(* Logix 5000 project; controller TFF vendor 1 type 14 code 107 rev 33.11; software revision 33.04; part 14 of 38 *)
(* tags used below, declared in another part *)
   ActionCode : DINT;   // Action Code
   ActionProperty : DINT;   // Action Property
   ActionStructure : DINT;   // Action Data Structure
   ActionTag : DINT;   // Action Tag
   ActionValue : REAL;   // Action Value
   Boolean : DINT;   // Boolean Operator
   Branch : BOOL;   // Conditional Branch Flag
   BranchStep : DINT;   // Branch Step Number
   BufferStep : DINT;   // Buffer Step
   Clear : BOOL;   // Clear Operation Table Flag
   Code : DINT;   // Global Code
   Criteria1BoolValue : BOOL;   // Criteria 1 Discrete Value
   Criteria1Code : DINT;   // Criteria 1 Code
   Criteria1Met : BOOL;   // Criteria 1 Met
   Criteria1Operator : DINT;   // Criteria 1 Operator
   Criteria1Property : DINT;   // Criteria 1 Property
   Criteria1RealValue : REAL;   // Criteria 1 Real Value
   Criteria1Structure : DINT;   // Criteria 1 Data Structure
   Criteria1Tag : DINT;   // Criteria 1 Tag
   Criteria1Type : BOOL;   // Criteria 1 Type 0=Real, 1=Boolean
   Criteria1Value : REAL;   // Criteria 1 Value
   Criteria2BoolValue : BOOL;   // Criteria 2 Discrete Value
   Criteria2Code : DINT;   // Criteria 2 Code
   Criteria2Met : BOOL;   // Criteria 2 Met
   Criteria2Operator : DINT;   // Criteria 2 Operator
   Criteria2Property : DINT;   // Criteria 2 Property
   Criteria2RealValue : REAL;   // Criteria 2 Real Value
   Criteria2Structure : DINT;   // Criteria 2 Data Structure
   Criteria2Tag : DINT;   // Criteria 2 Tag
   Criteria2Type : BOOL;   // Criteria 2 Type 0=Real, 1=Boolean
   Criteria2Value : REAL;   // Criteria 2 Value
   CriteriaMet : BOOL;   // Criteria Met
   DateTime : DINT[7];   // Date and Time
   ErrorCheck : BOOL;   // Error Check Flag
   Index : DINT;   // Index
   LastStep : DINT;   // Last Step
   NextStep : DINT;   // Next Step
   PendingStep : DINT;   // Current Step
   PhaseClear : BOOL;   // Phase Clear
   PhaseClearNumber : DINT;   // Phase Clear Number
   PhaseNumber : DINT;   // Phase FOR NEXT Index
   Pointer : DINT;   // Pointer
   PreRunLog : BOOL;   // Log Pre Run Set Points
   Property : DINT;   // Case Property
   Run : BOOL;   // Operation Run Status
   sAction : STRING10;   // Action Code String
   sActionProperty : STRING4;   // Action Property String
   sActionStructure : STRING4;   // Action Data Structure String
   sActionTag : STRING4;   // Action Tag String
   sBufferEvents : STRING50;   // Buffer Events String
   sCode : STRING10;   // Global code String
   sColon : STRING4;   // Colon separator String
   sComma : STRING4;   // Comma String
   sCriteria1 : STRING10;   // Criteria 1 Code String
   sCriteria1Property : STRING4;   // Criteria 1 Property String
   sCriteria1Structure : STRING4;   // Criteria 1 Data Structure String
   sCriteria1Tag : STRING4;   // Criteria 1 Tag String
   sCriteria2 : STRING10;   // Criteria 2 Code String
   sCriteria2Property : STRING4;   // Criteria 2 Property String
   sCriteria2Structure : STRING4;   // Criteria 2 Data Structure String
   sCriteria2Tag : STRING4;   // Criteria 2 Tag String
   sDateTime : STRING25;   // Date and Time String
   sPeriod : STRING4;   // Timer separator String
   sProperty : STRING4;   // Property String
   sStructure : STRING4;   // Structure String
   sTag : STRING4;   // Tag String
   sTemp : STRING50;   // Temp String
   Structure : DINT;   // Structure code
   sZero : STRING4;   // Zero String
   Tag : DINT;   // Tag value
   TempEvents : DINT;   // Temp Register
   TempSteps : DINT;
   Tenths : DINT;   // Thents (Date and Time management)
   ThisStep : DINT;   // This Step (Error management)
   Value : REAL;   // Temp Value
   AlarmAnalog : AlarmAnalog[50];   // Analog Alarm Array
   AlarmControl : AlarmControl;   // Alarm Control
   AlarmDeviation : AlarmDeviation[20];   // Control Loop Deviation Alarm Array
   AnalogPoint : AnalogInput[50];   // Analog Input Array
   BagInflate : BagInflate;
   CCPSystem : CCPSystem;   // CCP System Data
   ChartMark : ChartMark;   // Chart Mark
   Concentration : Concentration;
   ControlLoop : ControlLoop[20];   // Control Loop Array
   CPU_Scanning : BOOL;   // System Scanning Flag
   CriteriaFlag : CriteriaFlag;   // Criteria Flag used in CCP Recipe
   DerivedData : DerivedData;   // Derived data (user input and calculated values)
   Diafiltration : Diafiltration;
   DigitalPoint : DigitalPoint[150];   // Digital Point Array
   Drive : Drive[11];   // Drives Array
   Exchange_OUT : Exchange_OUT;   // Exchange Outputs
   ExternalTCU : BOOL;   // Use of External TCU
   ExternalWeight : BOOL;   // Use of External Weight
   FirstScanComplete : BOOL;   // First Scan Complete Flag
   FlowPath : FlowPath[64];   // Flow Path Array
   FQ_Conc : ALIAS FOR Totalizer[0];   // Concentration Totalizer
   FQ_Diaf : ALIAS FOR Totalizer[1];   // DiafiltrationTotalizer
   Gateway : Gateway;   // Gateway Control
   HoldTime : ALIAS FOR Timers[20];   // Hold Time
   LogVal : LoggedValue;   // Setpoints to be logged
   Membrane_Data : Membrane_Data;   // Membrane Data
   MiscBOOL : BOOL[64];   // Misc BOOL Values
   MiscDINT : DINT[32];   // Misc DINT Values
   MiscREAL : REAL[50];   // Misc Real Values
   Mixer : Mixer;   // Mixer config. structure
   Operation : Operation[6,251];   // Operation Table
   PCV101_Control : PCV_Control;   // PCV101 Control UDT
   PCV201_Control : PCV_Control;   // PCV201 Control UDT
   Phase : Phases[6];   // Phase Control Array
   Phase0 : ALIAS FOR Phase[0];   // Phase 0
   Phase0_Totalizer_Feed : ALIAS FOR PhaseTotalizer[0];   // Phase 0 Total Feed
   Phase0_Totalizer_Filtrate : ALIAS FOR PhaseTotalizer[6];   // Phase 0 Total Filtrate
   Phase0_Totalizer_Transfer : ALIAS FOR PhaseTotalizer[12];   // Phase 0 Total Transfer
   Phase1 : ALIAS FOR Phase[1];   // Phase 1
   Phase2 : ALIAS FOR Phase[2];   // Phase 2
   Phase3 : ALIAS FOR Phase[3];   // Phase 3
   Phase4 : ALIAS FOR Phase[4];   // Phase 4
   Phase5 : ALIAS FOR Phase[5];   // Phase 5
   PhaseTotalizer : PhaseTotalizer[18];   // Phase Totalizers Array
   PLCFault : FaultRecordType;   // PLC Major Fault Record
   ProcedureTime : ALIAS FOR Timers[19];   // Procedure Time
   Prompt : Prompt[7];   // Prompt Array
   Prompt0 : ALIAS FOR Prompt[0];   // Phase 0 Prompt
   Prompt1 : ALIAS FOR Prompt[1];   // Phase 1 Prompt
   Prompt2 : ALIAS FOR Prompt[2];   // Phase 2 Prompt
   Prompt3 : ALIAS FOR Prompt[3];   // Phase 3 Prompt
   Prompt4 : ALIAS FOR Prompt[4];   // Phase 4 Prompt
   Prompt5 : ALIAS FOR Prompt[5];   // Phase 5 Prompt
   SysControl : SysControl;   // General system status and command
   ThisSystem : SystemType;
   TIC101Control : TCUControl;
   TimerControl : TimerControl;   // Timer Control
   Timers : Timers[22];   // Timer Array
   Totalizer : Totalizers[20];   // Totalizers Array
   UserAlarm : UserAlarm;   // User Alarm (used in CCP Recipe)
   UserTotalizerManagement : UserTotalizerManagement;   // User Totalizer management
   Valve : Valve[100];   // Valve Array
   Y500A : ALIAS FOR DigitalOutput[10];
   Y500B : ALIAS FOR DigitalOutput[11];
   Y501A : ALIAS FOR DigitalOutput[12];
   Y501B : ALIAS FOR DigitalOutput[13];
   YA10 : ALIAS FOR DigitalPoint[59];
(* CCPSystem, continued *)

ROUTINE Branch   (* structured text *)
// Branch to Label Routine
   (* =======================================================================
   	Branch : Conditionnal branch management
   
   	List of treatments
   		- Get current action code
   		- Extract informations based on action code
   		- Jump to label and Jump Step processing
   
   -----------------------------------------------------------------------------------------------------------------------------------------------------
   	History
   		2019-DEC-24 - Merck - Q. Spindler - Initial version for Candidate Release 1.00.00.00.a
   =========================================================================*)
   
   
   (* Get current action code
   =========================================================================*)
   (*Get the pending step Action Code and Action Value from the operation array*)
   ActionCode := Operation[PhaseNumber,PendingStep].Action;
   ActionValue := Operation[PhaseNumber,PendingStep].ActionValue;
   
   (* Extract informations based on action code
   =========================================================================*)
   (*Extract the Structure, Tag and Property values from the action code. The action code is
   in the format SSTTTPP*)
   IF ActionCode <> 0 THEN;
   	DTOS (ActionCode, sAction);
   	IF sAction.LEN = 7 THEN;
   		MID (sAction, 2, 1, sActionStructure);
   		MID (sAction, 3, 3, sActionTag);
   		MID (sAction, 2, 6, sActionProperty);
   	ELSIF sAction.LEN = 6 THEN;
   		MID (sAction, 1, 1, sActionStructure);
   		MID (sAction, 3, 2, sActionTag);
   		MID (sAction, 2, 5, sActionProperty);
   	END_IF;
   	STOD (sActionStructure, ActionStructure);
   	STOD (sActionTag, ActionTag);
   	STOD (sActionProperty, ActionProperty);
   ELSE;
   	ActionStructure := 0;
   	ActionProperty := 0;
   END_IF;
   
   (* Jump to label and Jump Step processing
   =========================================================================*)
   (*Check to determine if action is a conditional branch, Structure=7 and Property=5*)
   BranchStep := 0;
   Phase[PhaseNumber].Label := 0;
   IF ActionStructure = 7 AND ActionProperty = 5  AND NOT Prompt[PhaseNumber].Pending THEN;
   	IF CriteriaMet THEN;
   		FOR BranchStep := 1 TO 250 DO;
   		(*If Jump to label action exist copy the label value in corresponding Phase label*)
   			IF Operation[PhaseNumber, BranchStep].Label = ActionValue THEN;
   				Phase[PhaseNumber].Label := ActionValue;
   				EXIT;
   			END_IF;
   		END_FOR;
   	ELSE;
   		(*Jump to BufferSteps routine and update Actual step number*)
   		JSR (BufferSteps);
   		Phase[PhaseNumber].ActualStep := (PendingStep + 1);
   	END_IF;
   
   ELSIF Phase[PhaseNumber].JumpPLC THEN;
   	FOR BranchStep := 1 TO 250 DO;
   		IF Operation[PhaseNumber, BranchStep].Step = Phase[PhaseNumber].JumpStep THEN;
   			Phase[PhaseNumber].ActualStep := BranchStep;
   			EXIT;
   		END_IF;
   	END_FOR;
   END_IF;
   
END_ROUTINE

ROUTINE BufferEvents   (* structured text *)
// Event Log Buffer Routine
   (* =======================================================================
   	Buffer Events : This routine scans all event code values defined in the event array downloaded by CCP6
   					If the value of the tag referenced by the code has changed from the last scan,the time stamp,
   					action code and new/old values are written to the buffer.
   					The buffer pointer used by CCP6 is updated after scanning all tags
   
   	Warning :		This code should not be modified without a control of change impact on the Recipe download check procedure of CCPRuntime.exe
   
   	List of treatments
   		- Get current action code
   		- Extract informations based on event code
   		- Navigate through the event categories
   		- Log Pre-run values
   		- Build event contents
   		- Reset flag and pointer
   
   -----------------------------------------------------------------------------------------------------------------------------------------------------
   	History
   		2019-DEC-24 - Merck - Q. Spindler - Initial version for Candidate Release 1.00.00.00.a
   		2020-MAR-30 - Merck - Q. Spindler - Modifications for Candidate Release 1.00.00.00.b
   					- Replace ActionProperty by Property for TIC
   					- Add SysControl.Zero_WI101_Cmd
   					- Add Valve.ZSOverride for valves limit switch alarms
   					- Add Gateway events
   		2020-SEP-18 - Merck - Q. Spindler - Modifications for Candidate Release 1.00.00.00.d
   					- Add ExternalWeight and ExternalTCU events
   		2022-JAN-21 - Merck - Q. Spindler - Modifications for Candidate Release 1.01.00.00.a
   					- Change resetting of sStructure in case of wrong code length by DTOS function
   		2022-SEP-21 - Actemium - J. Jaekel - Modifications for Candidate Release 1.01.00.01.a
   					- Add K and Q factor events
   =========================================================================*)
   
   
   (* Get the current pointer value
   =========================================================================*)
   STOD (CCPSystem.BufferEvents[0], Pointer);
   
   (* Extract informations based on event code
   =========================================================================*)
   (*Index through the event listing and get current value for each code*)
   (*The first element in the array is the array length*)
   FOR Index := 1 TO CCPSystem.EventList.Event[0] DO;
   
   	(*Extract the Structure, Tag and Property values from the code.  The code is in the format SSTTTPP*)
   	Code := CCPSystem.EventList.Event[Index];
   	DTOS (Code, sCode);
   
   		IF sCode.LEN = 7 THEN;
   			MID (sCode, 2, 1, sStructure);
   			MID (sCode, 3, 3, sTag);
   			MID (sCode, 2, 6, sProperty);
   		ELSIF sCode.LEN = 6 THEN;
   			MID (sCode, 1, 1, sStructure);
   			MID (sCode, 3, 2, sTag);
   			MID (sCode, 2, 5, sProperty);
   		ELSE;
   			(*Ignore if code length is not 6 or 7*)
   			DTOS (0, sStructure);
   		END_IF;
   		STOD (sStructure, Structure);
   		STOD (sTag, Tag);
   		STOD (sProperty, Property);
   
   	(* Tag:= 0; (*put in to handel error in congig files*)
   
   	Value := 0;
   
   (* Navigate through the event categories
   =========================================================================*)
   	(*Get the value based on the structure, tag and property*)
   	CASE	Structure OF
   		1: 	CASE	Property OF (*Analog Alarms*)
   			1:	IF AlarmAnalog[Tag].Override THEN Value := 1; ELSE Value := 0; END_IF;
   			2:	Value := AlarmAnalog[Tag].LOLO;
   			3:	Value := AlarmAnalog[Tag].LO;
   			4:	Value := AlarmAnalog[Tag].HI;
   			5:	Value := AlarmAnalog[Tag].HIHI;
   			6:	IF AlarmAnalog[Tag].LOLOAlarm THEN Value := 1; ELSE Value := 0; END_IF;
   			7:	IF AlarmAnalog[Tag].LOAlarm THEN Value := 1; ELSE Value := 0; END_IF;
   			8:	IF AlarmAnalog[Tag].HIAlarm THEN Value := 1; ELSE Value := 0; END_IF;
   			9:	IF AlarmAnalog[Tag].HIHIAlarm THEN Value := 1; ELSE Value := 0; END_IF;
   			END_CASE;
   		2: 	CASE	Property OF (*Deviation Alarms*)
   			1:	IF AlarmDeviation[Tag].Override THEN Value := 1; ELSE Value := 0; END_IF;
   			4:	Value := AlarmDeviation[Tag].HI;
   			5:	Value := AlarmDeviation[Tag].HIHI;
   			8:	IF AlarmDeviation[Tag].HIAlarm THEN Value := 1; ELSE Value := 0; END_IF;
   			9:	IF AlarmDeviation[Tag].HIHIAlarm THEN Value := 1; ELSE Value := 0; END_IF;
   			END_CASE;
   		3: 	CASE	Property OF (*Digital Alarms*)
   			1:	IF DigitalPoint[Tag].Override THEN Value := 1; ELSE Value := 0; END_IF;
   			6:	IF DigitalPoint[Tag].Alarm THEN Value := 1; ELSE Value := 0; END_IF;
   			7:	IF DigitalPoint[Tag].CurrentValue THEN Value := 1; ELSE Value := 0; END_IF;
   			END_CASE;
   		4: 	CASE	Property OF (*Analog Inputs*)
   			1:	Value := AnalogPoint[Tag].CurrentValue;
   			2:	Value := AnalogPoint[Tag].ScaledMin;
   			3:	Value := AnalogPoint[Tag].ScaledMax;
   			END_CASE;
   		5:	CASE	Property OF (*Control Loops*)
   			1:	IF ControlLoop[Tag].Manual THEN Value := 1; ELSE Value := 0; END_IF;
   			2:	IF ControlLoop[Tag].Auto1 THEN Value := 1; ELSE Value := 0; END_IF;
   			3:	IF ControlLoop[Tag].Auto2 THEN Value := 1; ELSE Value := 0; END_IF;
   			4:	IF ControlLoop[Tag].Auto3 THEN Value := 1; ELSE Value := 0; END_IF;
   			5:	IF ControlLoop[Tag].Auto4 THEN Value := 1; ELSE Value := 0; END_IF;
   			6:	Value := ControlLoop[Tag].SPManual;
   			7:	Value := ControlLoop[Tag].SPAuto1;
   			8:	Value := ControlLoop[Tag].SPAuto2;
   			9:	Value := ControlLoop[Tag].SPAuto3;
   			10:	Value := ControlLoop[Tag].SPAuto4;
   			11:	Value := ControlLoop[Tag].RampRate;
   			12:	Value := ControlLoop[Tag].Deadband;
   			13:	Value := ControlLoop[Tag].StableTime;
   			14:	Value := ControlLoop[Tag].KP[0];
   			15:	Value := ControlLoop[Tag].KI[0];
   			16:	Value := ControlLoop[Tag].KD[0];
   			17:	Value := ControlLoop[Tag].DB[0];
   			18:	Value := ControlLoop[Tag].KP[1];
   			19:	Value := ControlLoop[Tag].KI[1];
   			20:	Value := ControlLoop[Tag].KD[1];
   			21:	Value := ControlLoop[Tag].DB[1];
   			22:	Value := ControlLoop[Tag].KP[2];
   			23:	Value := ControlLoop[Tag].KI[2];
   			24:	Value := ControlLoop[Tag].KD[2];
   			25:	Value := ControlLoop[Tag].DB[2];
   			26:	IF ControlLoop[Tag].Stable THEN Value := 1; ELSE Value := 0; END_IF;
   			27:	IF ControlLoop[Tag].DBOK THEN Value := 1; ELSE Value := 0; END_IF;
   			28:	IF ControlLoop[Tag].RampStatus THEN Value := 1; ELSE Value := 0; END_IF;
   			END_CASE;
   		7:	CASE	Property OF (*Phase Control*)
   			1:	IF Phase[Tag].Run THEN Value := 1; ELSE Value := 0; END_IF;
   			2:	IF Phase[Tag].Stop THEN Value := 1; ELSE Value := 0; END_IF;
   			3:	IF Phase[Tag].Hold THEN Value := 1; ELSE Value := 0; END_IF;
   			4:	IF Phase[Tag].Pause THEN Value := 1; ELSE Value := 0; END_IF;
   			5:	IF Phase[Tag].Label = 0 THEN CCPSystem.EventList.Value[Index] := 0; END_IF; (*Ignore change to 0*)
   				Value := Phase[Tag].Label;
   			6:	IF Phase[Tag].JumpPLC THEN Value := 1; ELSE Value := 0; END_IF;
   			END_CASE;
   		8: 	CASE	Property OF (*Prompts*)
   			1:	IF Prompt[Tag].PromptOK THEN Value := 1; ELSE Value := 0; END_IF;
   			2:	IF Prompt[Tag].PromptYesNO THEN Value := 1; ELSE Value := 0; END_IF;
   			3:	IF Prompt[Tag].ResponseOK THEN Value := 1; ELSE Value := 0; END_IF;
   			4:	IF Prompt[Tag].ResponseYes THEN Value := 1; ELSE Value := 0; END_IF;
   			5:	IF Prompt[Tag].ResponseNo THEN Value := 1; ELSE Value := 0; END_IF;
   			END_CASE;
   		9: 	CASE	Property OF (*Pumps*)
   			1:	IF Drive[Tag].RunStatus THEN Value := 1; ELSE Value := 0; END_IF;
   			2:	IF Drive[Tag].Direction THEN Value := 1;ELSE Value := 0; END_IF;
   			3:	IF Drive[Tag].Mode THEN Value := 1; ELSE Value := 0; END_IF;
   			END_CASE;
   		10:	CASE	Property OF (*Exchange Output*)
   			1:	Value := Exchange_OUT.AO01;
   			2:	Value := Exchange_OUT.AO02;
   			3:	Value := Exchange_OUT.AO03;
   			4:	Value := Exchange_OUT.AO04;
   			5:	IF Exchange_OUT.DO01 THEN Value := 1; ELSE Value := 0; END_IF;
   			6:	IF Exchange_OUT.DO02 THEN Value := 1; ELSE Value := 0; END_IF;
   			7:	IF Exchange_OUT.DO03 THEN Value := 1; ELSE Value := 0; END_IF;
   			8:	IF Exchange_OUT.DO04 THEN Value := 1; ELSE Value := 0; END_IF;
   			9:	IF Exchange_OUT.DO05 THEN Value := 1; ELSE Value := 0; END_IF;
   			10:	IF Exchange_OUT.DO06 THEN Value := 1; ELSE Value := 0; END_IF;
   			11:	IF Exchange_OUT.DO07 THEN Value := 1; ELSE Value := 0; END_IF;
   			12:	IF Exchange_OUT.DO08 THEN Value := 1; ELSE Value := 0; END_IF;
   			END_CASE;
   		11:	CASE	Property OF (*Timers*)
   			3:	IF Timers[Tag].Enable THEN Value := 1; ELSE Value := 0; END_IF;
   			4:	IF Timers[Tag].Reset THEN Value := 1; ELSE Value := 0; END_IF;
   			END_CASE;
   		13:	CASE	Property OF (*Valves*)
   			2:	Value := Valve[Tag].StatusWord;
   			3:	IF Valve[Tag].Mode THEN Value := 1; ELSE Value := 0; END_IF;
   			4:	IF Valve[Tag].Alarm THEN Value := 1; ELSE Value := 0; END_IF;
   			5:	Value := Valve[Tag].Status;
   			6:	IF Valve[Tag].ZSOverride THEN Value := 1; ELSE Value := 0; END_IF;
   			END_CASE;
   		14:	CASE	Property OF (*Agitator*)
   			1:	IF Mixer.Mode THEN Value := 1; ELSE Value := 0; END_IF;
   			2:	Value := Mixer.SPManual;
   			3:	Value := Mixer.SPAutoMin;
   			4:	Value := Mixer.SPAutoMax;
   			5:	Value := Mixer.LevelMin;
   			6:	Value := Mixer.LevelMax;
   			END_CASE;
   		15:	CASE	Property OF (*Misc.*)
   			1:	IF MiscBOOL[Tag] THEN Value := 1; ELSE Value := 0; END_IF;
   			2:	Value := MiscDINT[Tag];
   			3:	Value := MiscREAL[Tag];
   			END_CASE;
   		16:	CASE	Property OF (*Alarm Control*)
   			1:	IF AlarmControl.EnableAllOut THEN Value := 1; ELSE Value := 0; END_IF;
   			2:	IF AlarmControl.DisableAllOut THEN Value := 1; ELSE Value := 0; END_IF;
   			3:	IF AlarmControl.AckOutput THEN Value := 1; ELSE Value := 0; END_IF;
   			6:	IF AlarmControl.EnableAllAnaSigOut THEN Value := 1; ELSE Value := 0; END_IF;
   			7:	IF AlarmControl.DisableAllAnaSigOut THEN Value := 1; ELSE Value := 0; END_IF;
   			END_CASE;
   		17:	CASE	Property OF (*Miscellaneous*)
   			1:	IF SysControl.DefaultOut THEN Value := 1; ELSE Value := 0; END_IF;
   			2:	IF ChartMark.Out THEN Value := 1; ELSE Value := 0; END_IF;
   			3:	IF SysControl.AllAutoOut THEN Value := 1; ELSE Value := 0; END_IF;
   			4:	IF UserTotalizerManagement.LogUserOut THEN Value := 1; ELSE Value := 0; END_IF;
   			5:	IF UserTotalizerManagement.StartUser THEN Value := 1; ELSE Value := 0; END_IF;
   			6:	IF UserTotalizerManagement.ResetUserOut THEN Value := 1; ELSE Value := 0; END_IF;
   			7:	IF SysControl.Tare_WI101_Cmd THEN Value := 1; ELSE Value := 0; END_IF;
   			8:	IF SysControl.ClearTare_WI101_Cmd THEN Value := 1; ELSE Value := 0; END_IF;
   			9:	IF SysControl.UV_Auto_Zero_Cmd THEN Value := 1; ELSE Value := 0; END_IF;
   			10:	IF SysControl.Zero_WI101_Cmd THEN Value := 1; ELSE Value := 0; END_IF;
   			11:	IF CCPSystem.DefaultOnComplete THEN Value := 1; ELSE Value := 0; END_IF;
   			12:	IF UserAlarm.NonCritical1 THEN Value := 1; ELSE Value := 0; END_IF;
   			13:	IF UserAlarm.Critical1 THEN Value := 1; ELSE Value := 0; END_IF;
   			14:	IF UserAlarm.NonCritical2 THEN Value := 1; ELSE Value := 0; END_IF;
   			15:	IF UserAlarm.Critical2 THEN Value := 1; ELSE Value := 0; END_IF;
   			16:	IF SysControl.Tare_PI001_Cmd THEN Value := 1; ELSE Value := 0; END_IF;
   			17:	IF SysControl.Tare_PI101_Cmd THEN Value := 1; ELSE Value := 0; END_IF;
   			18:	IF SysControl.Tare_PI201_Cmd THEN Value := 1; ELSE Value := 0; END_IF;
   			19:	IF SysControl.Tare_PI401_Cmd THEN Value := 1; ELSE Value := 0; END_IF;
   			20:	IF SysControl.Tare_PI601_Cmd THEN Value := 1; ELSE Value := 0; END_IF;
   			21:	IF BagInflate.cmd THEN Value := 1; ELSE Value := 0; END_IF;
   			22:	IF ExternalTCU THEN Value := 1; ELSE Value := 0; END_IF;
   			23:	IF ExternalWeight THEN Value := 1; ELSE Value := 0; END_IF;
   			END_CASE;
   		18:	CASE	Property OF (*Criteria Flag*)
   			1:	IF CriteriaFlag.Flag1 THEN Value := 1; ELSE Value := 0; END_IF;
   			2:	IF CriteriaFlag.Flag2 THEN Value := 1; ELSE Value := 0; END_IF;
   			3:	IF CriteriaFlag.Flag3 THEN Value := 1; ELSE Value := 0; END_IF;
   			4:	IF CriteriaFlag.Flag4 THEN Value := 1; ELSE Value := 0; END_IF;
   			5:	IF CriteriaFlag.Flag5 THEN Value := 1; ELSE Value := 0; END_IF;
   			END_CASE;
   		19:	CASE	Property OF (*Concentration*)
   			1:	IF FQ_Conc.Enable THEN Value := 1; ELSE Value := 0; END_IF;
   			2:	IF FQ_Conc.Reset THEN Value := 1; ELSE Value := 0; END_IF;
   			3:	IF Concentration.LogConcOut THEN Value := 1; ELSE Value := 0; END_IF;
   			4:	Value := Concentration.Conc_Init ;
   			5:	Value := Concentration.Conc_Final ;
   			6:	Value := Concentration.Conc_Final_Volume ;
   			7:	Value := DerivedData.HOLDUP ;
   			10: IF Concentration.Final_Conc_Volume_Reached THEN Value := 1; ELSE Value := 0; END_IF;
   			11: IF Concentration.Final_Conc_Protein_Reached THEN Value := 1; ELSE Value := 0; END_IF;
   			END_CASE;
   		20:	CASE	Property OF (*Diafiltration*)
   			1:	IF FQ_Diaf.Enable THEN Value := 1; ELSE Value := 0; END_IF;
   			2:	IF FQ_Diaf.Reset THEN Value := 1; ELSE Value := 0; END_IF;
   			3:	IF Diafiltration.LogDiafOut THEN Value := 1; ELSE Value := 0; END_IF;
   			4:	IF Diafiltration.Snap THEN Value := 1; ELSE Value := 0; END_IF;
   			5:	Value := Diafiltration.Diaf_Init ;
   			6:	Value := Diafiltration.Diaf_Final_Volume ;
   			10: IF Diafiltration.Final_Diaf_Volum_Reached THEN Value := 1; ELSE Value := 0; END_IF;
   			END_CASE;
   		21:	CASE	Property OF (*Membrane Data*)
   			1:	Value := Membrane_Data.Area ;
   			2:	Value := Membrane_Data.Density ;
   			3:	Value := DerivedData.FI101Q ;
   			4:	Value := DerivedData.FI201Q ;
   			5:	Value := DerivedData.FI401Q ;
   			6:	Value := DerivedData.FI101K ;
   			7:	Value := DerivedData.FI201K ;
   			8:	Value := DerivedData.FI401K ;
   			END_CASE;
   		22:	CASE	Property OF (*Gateway*)
   			1:	IF Tag <=31 THEN; (*Digital Actions*)
   					IF Gateway.RecipeAction_Digital[0].[Tag] THEN	Value := 1; ELSE Value := 0; END_IF;
   				ELSIF Tag <=63 THEN;
   					IF Gateway.RecipeAction_Digital[1].[Tag-32] THEN	Value := 1; ELSE Value := 0; END_IF;
   				END_IF;
   			2:	IF Tag <=19 THEN; (*Analog Actions*)
   				Value := Gateway.RecipeAction_Analog[Tag];
   				END_IF;
   			END_CASE;
   		23:	CASE	Property OF (*PCV Control*)
   			1:	IF PCV101_Control.FullOpen THEN Value := 1; ELSE Value := 0; END_IF;
   			2:	IF PCV101_Control.FullClose THEN Value := 1; ELSE Value := 0; END_IF;
   			3:	IF PCV201_Control.FullOpen THEN Value := 1; ELSE Value := 0; END_IF;
   			4:	IF PCV201_Control.FullClose THEN Value := 1; ELSE Value := 0; END_IF;
   			END_CASE;
   		24:	CASE	Property OF (*Event value.*)
   			1:	Value := LogVal.Value[Tag];
   			END_CASE;
   		25: CASE	Property OF (*Flow Paths*)
   			1:	IF FlowPath[Tag].Status THEN Value := 1; ELSE Value := 0; END_IF;
   			END_CASE;
   		26: CASE	Property OF (*Clamshell*)
   			1:	IF Y500A THEN Value := 1; ELSE Value := 0; END_IF;
   			2:	IF Y500B THEN Value := 1; ELSE Value := 0; END_IF;
   			3:	IF Y501A THEN Value := 1; ELSE Value := 0; END_IF;
   			4:	IF Y501B THEN Value := 1; ELSE Value := 0; END_IF;
   			11:  IF ThisSystem.MoldType = 123 THEN Value := 1; ELSE Value := 0; END_IF;
   			12:  IF ThisSystem.MoldType = 124 THEN Value := 1; ELSE Value := 0; END_IF;
   			13:  IF ThisSystem.MoldType = 126 THEN Value := 1; ELSE Value := 0; END_IF;
   			21:  IF ThisSystem.PreviousValue = 123 THEN Value := 1; ELSE Value := 0; END_IF;
   			22:  IF ThisSystem.PreviousValue = 124 THEN Value := 1; ELSE Value := 0; END_IF;
   			23:  IF ThisSystem.PreviousValue = 126 THEN Value := 1; ELSE Value := 0; END_IF;
   			END_CASE;
   		27:	CASE	Property OF (*TIC*)
   				1:	IF TIC101Control.RunCommand THEN Value := 1; ELSE Value := 0; END_IF;
   				2:  IF TIC101Control.Mode THEN Value := 1; ELSE Value := 0; END_IF;
   				3:	Value := TIC101Control.Offset;
   				4:	Value := TIC101Control.OffsetTime;
   				5:	Value := TIC101Control.LevelMin;
   			END_CASE;
   	(*Missing else statement accepted for the purpose of proper integration with CCPRuntime.exe*)
   	END_CASE;
   
   (* Log Pre-run values
   =========================================================================*)
   	(*Record value for Pre-Run Log if flag is set*)
   	IF PreRunLog THEN;
   		CCPSystem.EventList.PreRunValue[Index] := Value;
   	END_IF;
   
   
   (* Build event contents
   =========================================================================*)
   	(*Check for change in value*)
   	IF CCPSystem.EventList.Value[Index] <> Value THEN;
   		(*Increment pointer*)
   		Pointer := Pointer + 1;
   		(*Roll over pointer if equal to max*)
   		IF Pointer = 251 THEN Pointer := 1; END_IF;
   
   		(*Concatenate the action code to the date/time and add comma*)
   		DTOS (Code, sTemp);
   		CONCAT(sDateTime, sTemp, sBufferEvents);
   		CONCAT(sBufferEvents, sComma, sBufferEvents);
   
   		(*Concatenate the new value and add comma*)
   		RTOS (Value, sTemp);
   		CONCAT (sBufferEvents, sTemp, sBufferEvents);
   		CONCAT (sBufferEvents, sComma, sBufferEvents);
   
   		(*Concatenate the old value and store in the buffer*)
   		RTOS(CCPSystem.EventList.Value[Index], sTemp);
   		CONCAT(sBufferEvents, sTemp, CCPSystem.BufferEvents[Pointer]);
   
   		(*Clear the unused characters for null termination*)
   		TempEvents := CCPSystem.BufferEvents[Pointer].LEN;
   		WHILE TempEvents < 50 DO;
   			CCPSystem.BufferEvents[Pointer].DATA[TempEvents] := 0;
   			TempEvents := TempEvents + 1;
   		END_WHILE;
   
   		(*Save the new value for subsequent comparison*)
   		CCPSystem.EventList.Value[Index] := Value;
   	END_IF;
   END_FOR;
   
   (* Reset flag and pointer
   =========================================================================*)
   (*Clear the pre-run log flag*)
   PreRunLog := 0;
   
   (*Update the buffer pointer value after processing all events*)
   DTOS (Pointer, CCPSystem.BufferEvents[0]);
   
END_ROUTINE

ROUTINE BufferSteps   (* structured text *)
// Step Log Buffer Routine
   (* =======================================================================
   	Buffer Steps : This routine updates the step buffer when a step is executed
   
   	List of treatments
   		- Get current action code
   		- Compute the step value for the step buffer
   
   -----------------------------------------------------------------------------------------------------------------------------------------------------
   	History
   		2019-DEC-24 - Merck - Q. Spindler - Initial version for Candidate Release 1.00.00.00.a
   		2022-JAN-28 - Merck - Q. Spindler - Modifications for Candidate Release 1.01.00.00.a
   					- Limit LastStep to 0 minimum
   =========================================================================*)
   
   
   (* Get the current pointer value and increment
   =========================================================================*)
   STOD (CCPSystem.BufferSteps[0], Pointer);
   Pointer := Pointer + 1;
   (*Roll over pointer if equal to max*)
   IF Pointer = 251 THEN Pointer := 1; END_IF;
   DTOS (Pointer, CCPSystem.BufferSteps[0]);
   
   (* Compute the step value for the step buffer
   =========================================================================*)
   (*If the pending step number is the same as the last step number (named action list) then add 10000 to the buffer value*)
   LastStep := PendingStep - 1;
   IF LastStep < 0 THEN;
   	LastStep := 0;
   END_IF;
   IF Operation[PhaseNumber,PendingStep].Step = Operation[PhaseNumber,LastStep].Step THEN;
   	BufferStep := PhaseNumber * 1000 + (Operation[PhaseNumber,PendingStep].Step) + 10000;
   ELSE;
   	BufferStep := PhaseNumber * 1000 + (Operation[PhaseNumber,PendingStep].Step);
   END_IF;
   
   (*Convert the step value to a string and concatenate with the date/time*)
   DTOS (BufferStep, sTemp);
   CONCAT (sDateTime, sTemp, CCPSystem.BufferSteps[Pointer]);
   
   (*Clear the unused characters for null termination*)
   TempSteps := CCPSystem.BufferSteps[Pointer].LEN;
   WHILE TempSteps < 26 DO;
   	CCPSystem.BufferSteps[Pointer].DATA[TempSteps] := 0;
   	TempSteps := TempSteps + 1;
   END_WHILE;
END_ROUTINE

ROUTINE Clear   (* structured text *)
// Clear Operation Table
   (* =======================================================================
   	Clear : This routine loops through the entire operation array and clears
   			the step numbers, set Criteria1Value, Criteria2Value, ActionValue
   			to -999999.99 and sets all other values to -999.
   			This is executed at the start of each download.
   
   	List of treatments
   		- Initialize phase clear number
   		- Reset Operation data
   		- Reset Prompt messages
   		- In case of procedure RunAuto flag is set
   
   -----------------------------------------------------------------------------------------------------------------------------------------------------
   	History
   		2019-DEC-24 - Merck - Q. Spindler - Initial version for Candidate Release 1.00.00.00.a
   =========================================================================*)
   
   
   (* Initialize phase clear number
   =========================================================================*)
   (*One-Shot to set phase clear number to zero*)
   IF NOT PhaseClear THEN;
   	PhaseClearNumber := 0;
   	PhaseClear := 1;
   END_IF;
   
   (* Reset Operation data
   =========================================================================*)
   (*Step FOR-NEXT loop*)
   FOR PendingStep := 1 TO 250 DO;
   	Operation [PhaseClearNumber, PendingStep].Step := 0;
   	Operation [PhaseClearNumber, PendingStep].Criteria1 := -999;
   	Operation [PhaseClearNumber, PendingStep].Criteria1Operator := -999;
   	Operation [PhaseClearNumber, PendingStep].Boolean := -999;
   	Operation [PhaseClearNumber, PendingStep].Criteria2 := -999;
   	Operation [PhaseClearNumber, PendingStep].Criteria2Operator := -999;
   	Operation [PhaseClearNumber, PendingStep].Action := -999;
   	Operation [PhaseClearNumber, PendingStep].Label := -999;
   	Operation [PhaseClearNumber, PendingStep].Criteria1Value := -999999.99;
   	Operation [PhaseClearNumber, PendingStep].Criteria2Value := -999999.99;
   	Operation [PhaseClearNumber, PendingStep].ActionValue := -999999.99;
   END_FOR;
   
   PhaseClearNumber := PhaseClearNumber + 1;
   
   (* Reset Prompt messages
   =========================================================================*)
   IF PhaseClearNumber = 6 THEN;
   	(*Clear step buffer*)
   	CCPSystem.BufferSteps[0].LEN := 0;
   	(*State 11 ready for download*)
   	CCPSystem.State := 11;
   
   	Prompt0.PromptOK := 0;
   	Prompt0.PromptYesNO := 0;
   	Prompt1.PromptOK := 0;
   	Prompt1.PromptYesNO := 0;
   	Prompt2.PromptOK := 0;
   	Prompt2.PromptYesNO := 0;
   	Prompt3.PromptOK := 0;
   	Prompt3.PromptYesNO := 0;
   	Prompt4.PromptOK := 0;
   	Prompt4.PromptYesNO := 0;
   	Prompt5.PromptOK := 0;
   	Prompt5.PromptYesNO := 0;
   
   (* In case of procedure RunAuto flag is set
   =========================================================================*)
   	(*If part of a procedure then set the auto run flag so the operation will start when download is completed*)
   	IF CCPSystem.Procedure THEN;
   		CCPSystem.RunAuto := 1;
   	ELSE;
   		CCPSystem.RunAuto := 0;
   	END_IF;
   
   	PhaseClear := 0;
   
   END_IF;
   
END_ROUTINE

ROUTINE Complete   (* ladder *)
// Operation Complete Routine
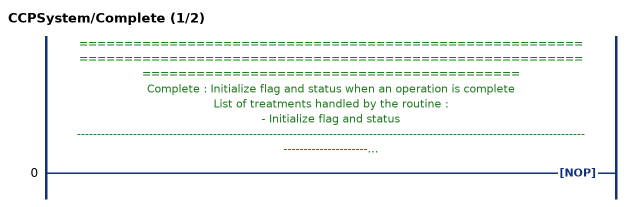
   // ==========================================================================================================================================================
   //                                                                                                Complete : Initialize flag and status when an operation is complete
   //                                                     List of treatments handled by the routine :
   //                                                          - Initialize flag and status
   //                                                     -----------------------------------------------------------------------------------------------------------------------------------------------------
   //                                                     History
   // 		2019-DEC-24 - Merck - Q. Spindler - Initial version for Candidate Release 1.00.00.00.a
   //                           2022-JAN-11 - Merck - Q. Spindler - Modifications for Candidate Release 1.01.00.00.a
   //                                 - Add unlatch of CCPSystem.Procedure when procedure is aborted
   // ========================================================================================================================================================
   0: NOP();
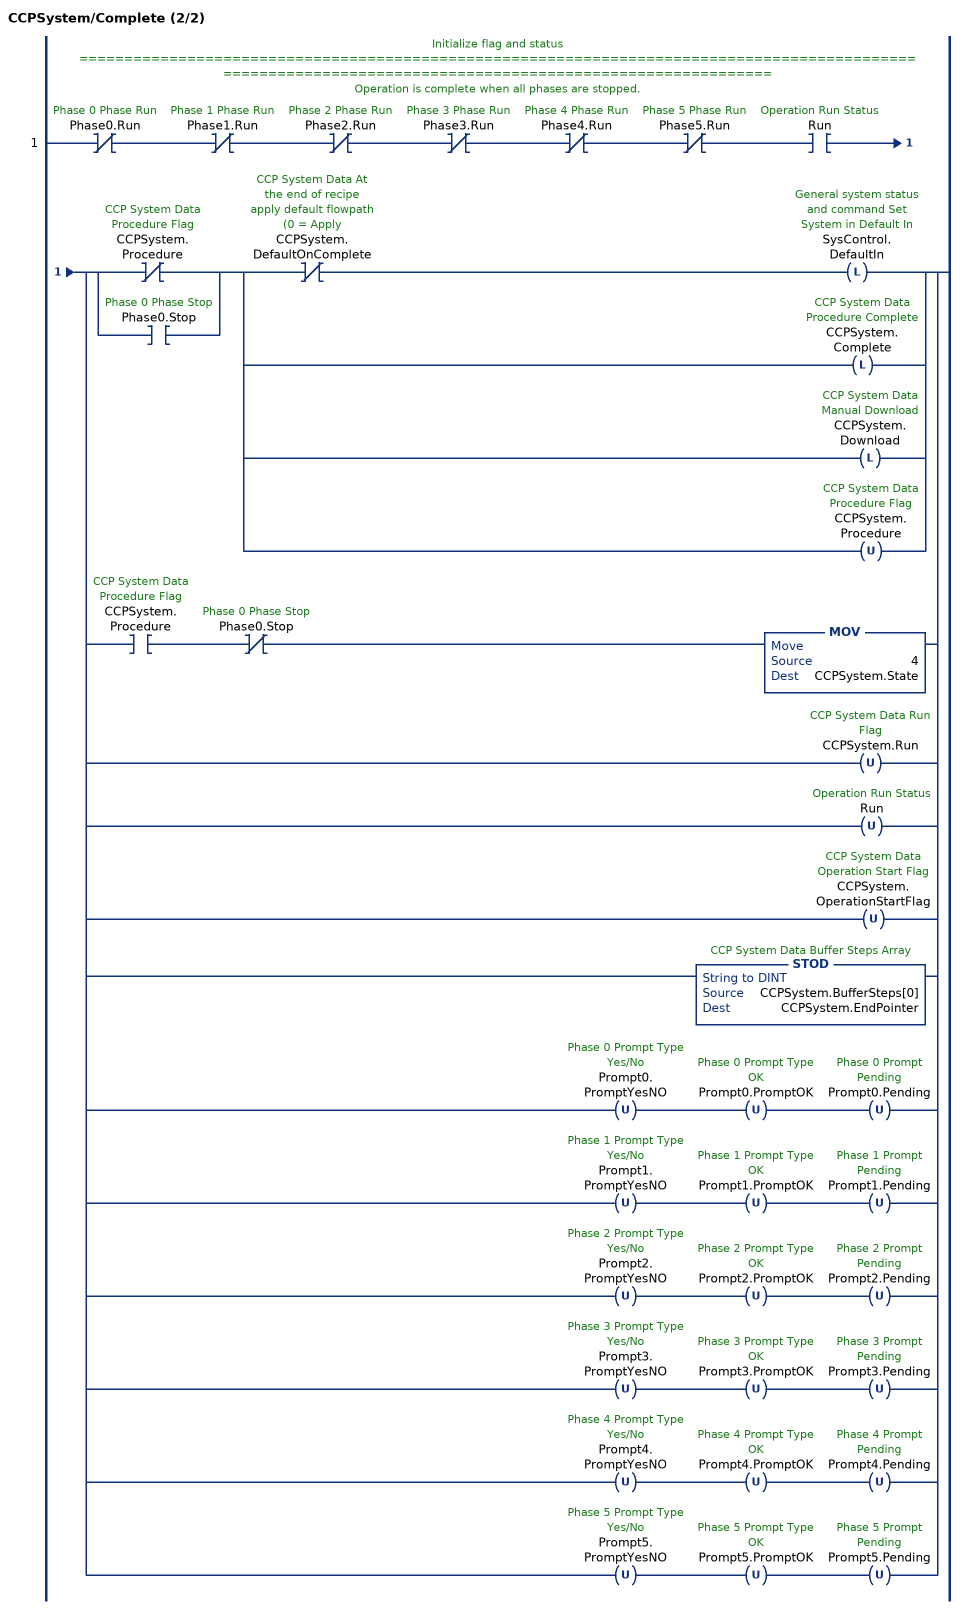
   // Initialize flag and status
   // ==========================================================================================================================================================
   // Operation is complete when all phases are stopped.
   1: XIO(Phase0.Run)XIO(Phase1.Run)XIO(Phase2.Run)XIO(Phase3.Run)XIO(Phase4.Run)XIO(Phase5.Run)XIC(Run)[[XIO(CCPSystem.Procedure) ,XIC(Phase0.Stop) ] [XIO(CCPSystem.DefaultOnComplete) OTL(SysControl.DefaultIn) ,OTL(CCPSystem.Complete) ,OTL(CCPSystem.Download) ,OTU(CCPSystem.Procedure) ] ,XIC(CCPSystem.Procedure) XIO(Phase0.Stop) MOV(4,CCPSystem.State) ,OTU(CCPSystem.Run) ,OTU(Run) ,OTU(CCPSystem.OperationStartFlag) ,STOD(CCPSystem.BufferSteps[0],CCPSystem.EndPointer) ,OTU(Prompt0.PromptYesNO) OTU(Prompt0.PromptOK) OTU(Prompt0.Pending) ,OTU(Prompt1.PromptYesNO) OTU(Prompt1.PromptOK) OTU(Prompt1.Pending) ,OTU(Prompt2.PromptYesNO) OTU(Prompt2.PromptOK) OTU(Prompt2.Pending) ,OTU(Prompt3.PromptYesNO) OTU(Prompt3.PromptOK) OTU(Prompt3.Pending) ,OTU(Prompt4.PromptYesNO) OTU(Prompt4.PromptOK) OTU(Prompt4.Pending) ,OTU(Prompt5.PromptYesNO) OTU(Prompt5.PromptOK) OTU(Prompt5.Pending) ];
END_ROUTINE

ROUTINE Criteria1   (* structured text *)
// Criteria 1 Routine
   (* =======================================================================
   	Criteria1 : Get the current criteria 1 code and verify if criteria met based on information extraction.
   				Update the criteria 1 bool and real value and the criteria type.
   
   	List of treatments
   		- Initialize Phase step number
   		- Extract informations based on criteria 1 code
   		- Navigate through the criteria categories and set Criteria bool and real value
   
   -----------------------------------------------------------------------------------------------------------------------------------------------------
   	History
   		2019-DEC-24 - Merck - Q. Spindler - Initial version for Candidate Release 1.00.00.00.a
   		2020-JUN-10 - Merck - Q. Spindler - Modifications for Candidate Release 1.00.00.00.c
   							- Remove CriteriaType for criteria VCF, DiaVolume,and CB.
   		2021-APR-22 - Merck - Q. Spindler - Modifications for Candidate Release 1.00.00.00.e
   							- Timers: Set the Time to 0 if the Reset flag is set to 1
   =========================================================================*)
   
   
   (* Initialize Phase step number
   =========================================================================*)
   (*If error check, pending step number is set by error check loop*)
   IF NOT ErrorCheck THEN;
   	PendingStep := Phase[PhaseNumber].ActualStep;
   	Phase[PhaseNumber].PendingStep := Operation[PhaseNumber,PendingStep].Step;
   	NextStep := PendingStep + 1;
   	IF PendingStep < 250 AND Operation[PhaseNumber,NextStep].Step <> 0 THEN;
   		Phase[PhaseNumber].NextStep := Operation[PhaseNumber,NextStep].Step;
   	ELSE;
   		Phase[PhaseNumber].NextStep := 0;
   	END_IF;
   END_IF;
   
   (* Extract informations based on criteria 1 code
   =========================================================================*)
   Criteria1Code := Operation[PhaseNumber,PendingStep].Criteria1;
   Criteria1Operator := Operation[PhaseNumber,PendingStep].Criteria1Operator;
   Criteria1Value := Operation[PhaseNumber,PendingStep].Criteria1Value;
   Boolean := Operation[PhaseNumber,PendingStep].Boolean;
   Criteria1Type := 0;
   
   (*Extract the Structure, Tag and Property values from the criteria code.  The criteria code is
   in the format SSTTTPP*)
   
   IF Criteria1Code <> 0 THEN;
   	DTOS (Criteria1Code, sCriteria1);
   	IF sCriteria1.LEN = 7 THEN;
   		MID (sCriteria1, 2, 1, sCriteria1Structure);
   		MID (sCriteria1, 3, 3, sCriteria1Tag);
   		MID (sCriteria1, 2, 6, sCriteria1Property);
   	ELSIF sCriteria1.LEN = 6 THEN;
   		MID (sCriteria1, 1, 1, sCriteria1Structure);
   		MID (sCriteria1, 3, 2, sCriteria1Tag);
   		MID (sCriteria1, 2, 5, sCriteria1Property);
   	ELSE;
   		CCPSystem.Error := 2;
   	END_IF;
   	STOD (sCriteria1Structure, Criteria1Structure);
   	STOD (sCriteria1Tag, Criteria1Tag);
   	STOD (sCriteria1Property, Criteria1Property);
   ELSE;
   	Criteria1Structure := 0;
   END_IF;
   
   (* Navigate through the criteria categories and set Criteria bool and real value
   =========================================================================*)
   CASE	Criteria1Structure OF
   	0:	; (*No Criteria*)
   	3:	CASE	Criteria1Property OF (*Digital Points*)
   			1:	Criteria1BoolValue := DigitalPoint[Criteria1Tag].CurrentValue;
   				Criteria1Type := 1;
   			2:	Criteria1BoolValue := DigitalPoint[Criteria1Tag].Alarm;
   				Criteria1Type := 1;
   			3:	Criteria1BoolValue := DigitalPoint[Criteria1Tag].SoftInput;
   				Criteria1Type := 1;
   		ELSE 	CCPSystem.Error := 2;
   		END_CASE;
   	4: 	CASE	Criteria1Property OF (*Analog Inputs*)
   			1:	Criteria1RealValue := AnalogPoint[Criteria1Tag].CurrentValue;
   		ELSE 	CCPSystem.Error := 2;
   		END_CASE;
   	5:	CASE	Criteria1Property OF (*Control Loops*)
   			18:	Criteria1BoolValue := ControlLoop[Criteria1Tag].Stable;
   				Criteria1Type := 1;
   			19:	Criteria1BoolValue := ControlLoop[Criteria1Tag].DBOK;
   				Criteria1Type := 1;
   			20:	Criteria1BoolValue := ControlLoop[Criteria1Tag].RampStatus;
   				Criteria1Type := 1;
   		ELSE 	CCPSystem.Error := 2;
   		END_CASE;
   	7:	CASE	Criteria1Property OF (*Phase Control*)
   			1:	Criteria1BoolValue := Phase[Criteria1Tag].Run;
   				Criteria1Type := 1;
   			3:	Criteria1BoolValue := Phase[Criteria1Tag].Hold;
   				Criteria1Type := 1;
   			4:	Criteria1BoolValue := Phase[Criteria1Tag].Pause;
   		ELSE 	CCPSystem.Error := 2;
   		END_CASE;
   	8: 	CASE	Criteria1Property OF (*Prompts*)
   			3:	Criteria1BoolValue := Prompt[PhaseNumber].ResponseOK;
   				Criteria1Type := 1;
   			4:	Criteria1BoolValue := Prompt[PhaseNumber].ResponseYes;
   				Criteria1Type := 1;
   			5:	Criteria1BoolValue := Prompt[PhaseNumber].ResponseNo;
   				Criteria1Type := 1;
   		ELSE 	CCPSystem.Error := 2;
   		END_CASE;
   	9: 	CASE	Criteria1Property OF (*Pumps*)
   			2:	Criteria1BoolValue := Drive[Criteria1Tag].RunStatus;
   				Criteria1Type := 1;
   		ELSE 	CCPSystem.Error := 2;
   		END_CASE;
   	11:	CASE	Criteria1Property OF (*Timers*)
   			1:	IF Timers[Criteria1Tag].Reset THEN Criteria1RealValue := 0;
   				ELSE Criteria1RealValue := Timers[Criteria1Tag].TotalSeconds; (*Total Time*) END_IF;
   			2:	Criteria1Tag := Criteria1Tag + PhaseNumber; (*Add phase number to address correct step timer*)
   				IF Timers[Criteria1Tag].Reset THEN Criteria1RealValue := 0;
   				ELSE Criteria1RealValue := Timers[Criteria1Tag].TotalSeconds; (*Step Time*) END_IF;
   		ELSE 	CCPSystem.Error := 2;
   		END_CASE;
   	12:	CASE	Criteria1Property OF (*Totalizers*)
   			1:	Criteria1RealValue := PhaseTotalizer[Criteria1Tag].Phase;
   			2:	Criteria1Tag := Criteria1Tag + PhaseNumber; (*Add phase number to address correct step totalizer*)
   				Criteria1RealValue := PhaseTotalizer[Criteria1Tag].Step;
   			3:	Criteria1RealValue := PhaseTotalizer[Criteria1Tag].Pause;
   			4:	Criteria1RealValue := PhaseTotalizer[Criteria1Tag].User;
   			5:	Criteria1RealValue := PhaseTotalizer[Criteria1Tag].Procedure;
   			8:	Criteria1RealValue := Totalizer[Criteria1Tag].Total;
   		ELSE 	CCPSystem.Error := 2;
   		END_CASE;
   	13:	CASE	Criteria1Property OF (*Valves*)
   			2:	Criteria1RealValue := Valve[Criteria1Tag].StatusWord;
   		ELSE 	CCPSystem.Error := 2;
   		END_CASE;
   	15:	CASE	Criteria1Property OF (*Misc.*)
   			1:	Criteria1BoolValue := MiscBOOL[Criteria1Tag];
   				Criteria1Type := 1;
   			2:	Criteria1RealValue := MiscDINT[Criteria1Tag];
   			3:	Criteria1RealValue := MiscREAL[Criteria1Tag];
   		ELSE 	CCPSystem.Error := 2;
   		END_CASE;
   	17:	CASE	Criteria1Property OF (*Miscellaneous*)
   			11:	Criteria1BoolValue := CCPSystem.DefaultOnComplete ;
   				Criteria1Type := 1;
   		ELSE 	CCPSystem.Error := 2;
   		END_CASE;
   	18:	CASE	Criteria1Property OF (*Criteria Flag*)
   			1:	Criteria1BoolValue := CriteriaFlag.Flag1 ;
   				Criteria1Type := 1;
   			2:	Criteria1BoolValue := CriteriaFlag.Flag2 ;
   				Criteria1Type := 1;
   			3:	Criteria1BoolValue := CriteriaFlag.Flag3 ;
   				Criteria1Type := 1;
   			4:	Criteria1BoolValue := CriteriaFlag.Flag4 ;
   				Criteria1Type := 1;
   			5:	Criteria1BoolValue := CriteriaFlag.Flag5 ;
   				Criteria1Type := 1;
   		ELSE 	CCPSystem.Error := 2;
   		END_CASE;
   	19:	CASE	Criteria1Property OF (*Concentration*)
   			1:	Criteria1RealValue := Concentration.VCF;
   			2:	Criteria1RealValue := Concentration.CB;
   			3:	Criteria1BoolValue := Concentration.Final_Conc_Volume_Reached ;
   				Criteria1Type := 1;
   			4:	Criteria1BoolValue := Concentration.Final_Conc_Protein_Reached ;
   				Criteria1Type := 1;
   		ELSE 	CCPSystem.Error := 2;
   		END_CASE;
   	20:	CASE	Criteria1Property OF (*Diafiltration*)
   			1:	Criteria1RealValue := Diafiltration.Diaf_Volume;
   			2:	Criteria1BoolValue := Diafiltration.Final_Diaf_Volum_Reached ;
   				Criteria1Type := 1;
   		ELSE 	CCPSystem.Error := 2;
   		END_CASE;
   	22:	CASE	Criteria1Property OF (*Gateway*)
   			(*Digital*)
   			1:	IF Criteria1Tag <=31 THEN;
   					Criteria1BoolValue := Gateway.RecipeCriteria_Digital[0].[Criteria1Tag];
   				ELSIF Criteria1Tag <=63 THEN;
   					Criteria1BoolValue := Gateway.RecipeCriteria_Digital[1].[Criteria1Tag-32];
   				END_IF;
   				Criteria1Type := 1;
   			(*Analog*)
   			2:	Criteria1RealValue := Gateway.RecipeCriteria_Analog[Criteria1Tag];
   		ELSE 	CCPSystem.Error := 2;
   		END_CASE;
   	25: CASE	Criteria1Property OF (*Flow Paths*)
   			2:	Criteria1BoolValue := FlowPath[Criteria1Tag].Status;
   				Criteria1Type := 1;
   		ELSE 	CCPSystem.Error := 2;
   		END_CASE;
   ELSE	CCPSystem.Error := 2;
   END_CASE;
   
END_ROUTINE

ROUTINE Criteria2   (* structured text *)
// Criteria 2 Routine
   (* =======================================================================
   	Criteria2 : Get the current criteria 2 code and verify if criteria met based on information extraction.
   				Update the criteria 2 bool and real value and the criteria type.
   
   	List of treatments
   		- Initialize Phase step number
   		- Extract informations based on criteria 2 code
   		- Navigate through the criteria categories and set Criteria bool and real value
   
   -----------------------------------------------------------------------------------------------------------------------------------------------------
   	History
   		2019-DEC-24 - Merck - Q. Spindler - Initial version for Candidate Release 1.00.00.00.a
   		2020-JUN-10 - Merck - Q. Spindler - Modifications for Candidate Release 1.00.00.00.c
   							- Remove CriteriaType for criteria VCF, DiaVolume,and CB.
   		2021-APR-22 - Merck - Q. Spindler - Modifications for Candidate Release 1.00.00.00.e
   							- Timers: Set the Time to 0 if the Reset flag is set to 1
   =========================================================================*)
   
   (* Extract informations based on criteria 2 code
   =========================================================================*)
   Criteria2Code := Operation[PhaseNumber,PendingStep].Criteria2;
   Criteria2Operator := Operation[PhaseNumber,PendingStep].Criteria2Operator;
   Criteria2Value := Operation[PhaseNumber,PendingStep].Criteria2Value;
   Criteria2Type := 0;
   
   IF Criteria2Code <> 0 THEN;
   	DTOS (Criteria2Code, sCriteria2);
   	IF sCriteria2.LEN = 7 THEN;
   		MID (sCriteria2, 2, 1, sCriteria2Structure);
   		MID (sCriteria2, 3, 3, sCriteria2Tag);
   		MID (sCriteria2, 2, 6, sCriteria2Property);
   	ELSIF sCriteria2.LEN = 6 THEN;
   		MID (sCriteria2, 1, 1, sCriteria2Structure);
   		MID (sCriteria2, 3, 2, sCriteria2Tag);
   		MID (sCriteria2, 2, 5, sCriteria2Property);
   	ELSE;
   		CCPSystem.Error := 5;
   	END_IF;
   	STOD (sCriteria2Structure, Criteria2Structure);
   	STOD (sCriteria2Tag, Criteria2Tag);
   	STOD (sCriteria2Property, Criteria2Property);
   ELSE;
   	Criteria2Structure := 0;
   END_IF;
   
   (* Navigate through the criteria categories and set Criteria bool and real value
   =========================================================================*)
   CASE	Criteria2Structure OF
   	0:	; (*No Criteria*)
   	3:	CASE	Criteria2Property OF (*Digital Points*)
   			1:	Criteria2BoolValue := DigitalPoint[Criteria2Tag].CurrentValue;
   				Criteria2Type := 1;
   			2:	Criteria2BoolValue := DigitalPoint[Criteria2Tag].Alarm;
   				Criteria2Type := 1;
   			3:	Criteria2BoolValue := DigitalPoint[Criteria2Tag].SoftInput;
   				Criteria2Type := 1;
   		ELSE 	CCPSystem.Error := 2;
   		END_CASE;
   	4: 	CASE	Criteria2Property OF (*Analog Inputs*)
   			1:	Criteria2RealValue := AnalogPoint[Criteria2Tag].CurrentValue;
   		ELSE 	CCPSystem.Error := 5;
   		END_CASE;
   	5:	CASE	Criteria2Property OF (*Control Loops*)
   			18:	Criteria2BoolValue := ControlLoop[Criteria2Tag].Stable;
   				Criteria2Type := 1;
   			19:	Criteria2BoolValue := ControlLoop[Criteria2Tag].DBOK;
   				Criteria2Type := 1;
   			20:	Criteria2BoolValue := ControlLoop[Criteria2Tag].RampStatus;
   				Criteria2Type := 1;
   		ELSE 	CCPSystem.Error := 5;
   		END_CASE;
   	7:	CASE	Criteria2Property OF (*Phase Control*)
   			1:	Criteria2BoolValue := Phase[Criteria2Tag].Run;
   				Criteria2Type := 1;
   			3:	Criteria2BoolValue := Phase[Criteria2Tag].Hold;
   				Criteria2Type := 1;
   			4:	Criteria2BoolValue := Phase[Criteria2Tag].Pause;
   			6:	Criteria2Tag := Criteria2Tag + PhaseNumber;
   				Criteria2RealValue := Phase[Criteria2Tag].Crit1MetTime;
   		ELSE 	CCPSystem.Error := 5;
   		END_CASE;
   	8: 	CASE	Criteria2Property OF (*Prompts*)
   			3:	Criteria2BoolValue := Prompt[PhaseNumber].ResponseOK;
   				Criteria2Type := 1;
   			4:	Criteria2BoolValue := Prompt[PhaseNumber].ResponseYes;
   				Criteria2Type := 1;
   			5:	Criteria2BoolValue := Prompt[PhaseNumber].ResponseNo;
   				Criteria2Type := 1;
   		ELSE 	CCPSystem.Error := 5;
   		END_CASE;
   	9: 	CASE	Criteria2Property OF (*Pumps*)
   			2:	Criteria2BoolValue := Drive[Criteria2Tag].RunStatus;
   				Criteria2Type := 1;
   		ELSE 	CCPSystem.Error := 5;
   		END_CASE;
   	11:	CASE	Criteria2Property OF (*Timers*)
   			1:	IF Timers[Criteria2Tag].Reset THEN Criteria2RealValue := 0;
   				ELSE Criteria2RealValue := Timers[Criteria2Tag].TotalSeconds; (*Total Time*) END_IF;
   			2:	Criteria2Tag := Criteria2Tag + PhaseNumber; (*Add phase number to address correct step timer*)
   				IF Timers[Criteria2Tag].Reset THEN Criteria2RealValue := 0;
   				ELSE Criteria2RealValue := Timers[Criteria2Tag].TotalSeconds; (*Step Time*) END_IF;
   		ELSE 	CCPSystem.Error := 5;
   		END_CASE;
   	12:	CASE	Criteria2Property OF (*Totalizers*)
   			1:	Criteria2RealValue := PhaseTotalizer[Criteria2Tag].Phase;
   			2:	Criteria2Tag := Criteria2Tag + PhaseNumber; (*Add phase number to address correct step totalizer*)
   				Criteria2RealValue := PhaseTotalizer[Criteria2Tag].Step;
   			3:	Criteria2RealValue := PhaseTotalizer[Criteria2Tag].Pause;
   			4:	Criteria2RealValue := PhaseTotalizer[Criteria2Tag].User;
   			5:	Criteria2RealValue := PhaseTotalizer[Criteria2Tag].Procedure;
   			8:	Criteria2RealValue := Totalizer[Criteria2Tag].Total;
   		ELSE 	CCPSystem.Error := 5;
   		END_CASE;
   	13:	CASE	Criteria2Property OF (*Valves*)
   			2:	Criteria2RealValue := Valve[Criteria2Tag].StatusWord;
   		ELSE 	CCPSystem.Error := 5;
   		END_CASE;
   	15:	CASE	Criteria2Property OF (*Misc.*)
   			1:	Criteria2BoolValue := MiscBOOL[Criteria2Tag];
   				Criteria2Type := 1;
   			2:	Criteria2RealValue := MiscDINT[Criteria2Tag];
   			3:	Criteria2RealValue := MiscREAL[Criteria2Tag];
   		ELSE 	CCPSystem.Error := 5;
   		END_CASE;
   	17:	CASE	Criteria2Property OF (*Miscellaneous*)
   			11:	Criteria2BoolValue := CCPSystem.DefaultOnComplete ;
   				Criteria2Type := 1;
   		ELSE 	CCPSystem.Error := 5;
   		END_CASE;
   	18:	CASE	Criteria2Property OF (*Criteria Flag*)
   			1:	Criteria2BoolValue := CriteriaFlag.Flag1 ;
   				Criteria2Type := 1;
   			2:	Criteria2BoolValue := CriteriaFlag.Flag2 ;
   				Criteria2Type := 1;
   			3:	Criteria2BoolValue := CriteriaFlag.Flag3 ;
   				Criteria2Type := 1;
   			4:	Criteria2BoolValue := CriteriaFlag.Flag4 ;
   				Criteria2Type := 1;
   			5:	Criteria2BoolValue := CriteriaFlag.Flag5 ;
   				Criteria2Type := 1;
   		ELSE 	CCPSystem.Error := 5;
   		END_CASE;
   	19:	CASE	Criteria2Property OF (*Concentration*)
   			1:	Criteria2RealValue := Concentration.VCF;
   			2:	Criteria2RealValue := Concentration.CB;
   			3:	Criteria2BoolValue := Concentration.Final_Conc_Volume_Reached ;
   				Criteria2Type := 1;
   			4:	Criteria2BoolValue := Concentration.Final_Conc_Protein_Reached ;
   				Criteria2Type := 1;
   		ELSE 	CCPSystem.Error := 5;
   		END_CASE;
   	20:	CASE	Criteria2Property OF (*Diafiltration*)
   			1:	Criteria2RealValue := Diafiltration.Diaf_Volume;
   			2:	Criteria2BoolValue := Diafiltration.Final_Diaf_Volum_Reached ;
   				Criteria2Type := 1;
   		ELSE 	CCPSystem.Error := 5;
   		END_CASE;
   	22:	CASE	Criteria2Property OF (*Gateway*)
   			(*Digital*)
   			1:	IF Criteria2Tag <=31 THEN;
   					Criteria2BoolValue := Gateway.RecipeCriteria_Digital[0].[Criteria2Tag];
   				ELSIF Criteria2Tag <=63 THEN;
   					Criteria2BoolValue := Gateway.RecipeCriteria_Digital[1].[Criteria2Tag-32];
   				END_IF;
   				Criteria2Type := 1;
   			(*Analog*)
   			2:	Criteria2RealValue := Gateway.RecipeCriteria_Analog[Criteria2Tag];
   		ELSE 	CCPSystem.Error := 5;
   		END_CASE;
   	25: 	CASE	Criteria2Property OF (*Flow Paths*)
   			2:	Criteria2BoolValue := FlowPath[Criteria2Tag].Status;
   				Criteria2Type := 1;
   		ELSE 	CCPSystem.Error := 5;
   		END_CASE;
   ELSE	CCPSystem.Error := 5;
   END_CASE;
   
END_ROUTINE

ROUTINE DateTime   (* structured text *)
// System Date and Time Routine
   (* =======================================================================
   	DateTime : 	This routine returns a string value of date and time in the format "MMDDYYYY,HH:MM:SS.x,".
   				The result is stored in the program tag sDateTime.
   				This string will be used by the BufferEvents and BufferSteps routines for time stamping.
   
   	List of treatments
   		- Get system date and time with GSV instruction
   		- Convert the date and time in DINT format to string format
   
   -----------------------------------------------------------------------------------------------------------------------------------------------------
   	History
   		2019-DEC-24 - Merck - Q. Spindler - Initial version for Candidate Release 1.00.00.00.a
   =========================================================================*)
   
   
   (* Get system date and time with GSV instruction
   =========================================================================*)
   
   (*Get the current date and time from the processor*)
   (*The date and time are stored in an array of 7 values*)
   	GSV (WALLCLOCKTIME, , DateTime, DateTime[0]);
   
   (* Convert the date and time in DINT format to string format
   =========================================================================*)
   (*Month*)
   	DTOS (DateTime[1], sDateTime);
   	(*Add leading zero if value is 1 character*)
   	IF sDateTime.LEN = 1 Then;
   		CONCAT (sZero, sDateTime, sDateTime);
   	END_IF;
   (*Day*)
   	DTOS (DateTime[2], sTemp);
   	(*Add leading zero if value is 1 character*)
   	IF sTemp.LEN = 1 Then;
   		CONCAT (sZero, sTemp, sTemp);
   	END_IF;
   	CONCAT (sDateTime, sTemp, sDateTime);
   (*Year*)
   	DTOS (DateTime[0], sTemp);
   	CONCAT (sDateTime, sTemp, sDateTime);
   	CONCAT (sDateTime, sComma, sDateTime);
   (*Hours*)
   	DTOS (DateTime[3], sTemp);
   	(*Add leading zero if value is 1 character*)
   	IF sTemp.LEN = 1 Then;
   		CONCAT (sZero, sTemp, sTemp);
   	END_IF;
   	CONCAT (sDateTime, sTemp, sDateTime);
   	CONCAT (sDateTime, sColon, sDateTime);
   (*Minutes*)
   	DTOS (DateTime[4], sTemp);
   	(*Add leading zero if value is 1 character*)
   	IF sTemp.LEN = 1 Then;
   		CONCAT (sZero, sTemp, sTemp);
   	END_IF;
   	CONCAT (sDateTime, sTemp, sDateTime);
   	CONCAT (sDateTime, sColon, sDateTime);
   (*Seconds*)
   	DTOS (DateTime[5], sTemp);
   	(*Add leading zero if value is 1 character*)
   	IF sTemp.LEN = 1 Then;
   		CONCAT (sZero, sTemp, sTemp);
   	END_IF;
   	CONCAT (sDateTime, sTemp, sDateTime);
   	CONCAT (sDateTime, sPeriod, sDateTime);
   (*Tenth Seconds*)
   	(*Round the microseconds value to tenths seconds*)
   	Tenths := DateTime[6] / 100000;
   	DTOS (Tenths, sTemp);
   	CONCAT (sDateTime, sTemp, sDateTime);
   	CONCAT (sDateTime, sComma, sDateTime);
   
END_ROUTINE

ROUTINE Error   (* structured text *)
// Step Error Checking
   (* =======================================================================
   	Error : This routine loops through all steps of one phase per processor scan to detect an error
   
   	List of treatments
   		- Initialize
   		- Error check processing
   		- Error found
   		- No error found
   
   -----------------------------------------------------------------------------------------------------------------------------------------------------
   	History
   		2019-DEC-24 - Merck - Q. Spindler - Initial version for Candidate Release 1.00.00.00.a
   =========================================================================*)
   
   
   (* Initialize
   =========================================================================*)
   (*Initialize error check values first time*)
   IF NOT ErrorCheck THEN;
   	CCPSystem.Error := 0;
   	CCPSystem.ErrorStep:= 0;
   	CCPSystem.ErrorPhase := 0;
   	PhaseNumber := 0;
   	ErrorCheck := 1;
   ELSE;
   	PhaseNumber := PhaseNumber + 1;
   END_IF;
   (* PhaseNumber := 5;*)
   (*Reset the total and last step values*)
   Phase[PhaseNumber].TotalSteps := 0;
   LastStep := 0;
   
   (* Error check processing
   =========================================================================*)
   (*Loop through the steps.  If step number is zero, complete*)
   FOR PendingStep := 1 TO 250 DO;
   	IF Operation[PhaseNumber, PendingStep].Step = 0 THEN;
   		EXIT;
   	END_IF;
   
   	(*Step Number Error Check*)
   	(*Verify step number is equal to or one greater than the previous step number*)
   	ThisStep := Operation[PhaseNumber, PendingStep].Step;
   	IF ThisStep <> LastStep + 1 AND ThisStep <> LastStep THEN;
   		CCPSystem.Error := 1;
   		EXIT;
   	END_IF;
   	LastStep := ThisStep;
   	Phase[PhaseNumber].TotalSteps := PendingStep;
   
   	(*Criteria 1 Error Check*)
   	JSR (Criteria1);
   	IF CCPSystem.Error <> 0 THEN;
   		EXIT;
   	END_IF;
   	IF Criteria1Operator <> 0 AND Criteria1Operator <> 1 AND Criteria1Operator <> 2 AND Criteria1Operator <> 4 THEN;
   		CCPSystem.Error := 3;
   		EXIT;
   	ELSIF Boolean > 2 THEN;
   		CCPSystem.Error := 4;
   		EXIT;
   	ELSIF Criteria1Value = -999999.99 THEN;
   		CCPSystem.Error := 9;
   		EXIT;
   	END_IF;
   
   	(*Criteria 2 Error Check*)
   	JSR (Criteria2);
   	IF CCPSystem.Error <> 0 THEN;
   		EXIT;
   	END_IF;
   	IF Criteria2Operator <> 0 AND Criteria2Operator <> 1 AND Criteria2Operator <> 2 AND Criteria2Operator <> 4 THEN;
   		CCPSystem.Error := 6;
   		EXIT;
   	ELSIF Criteria2Value = -999999.99 THEN;
   		CCPSystem.Error := 10;
   		EXIT;
   	END_IF;
   
   	(*Action Error Check*)
   	JSR (Action);
   	IF CCPSystem.Error <> 0 THEN;
   		EXIT;
   	END_IF;
   	IF ActionValue = -999999.99 THEN;
   		CCPSystem.Error := 11;
   		EXIT;
   	END_IF;
   
   	(*Label Error Check*)
   	IF  Operation[PhaseNumber, PendingStep].Label > 20 THEN;
   		CCPSystem.Error := 8;
   		EXIT;
   	END_IF;
   END_FOR;
   
   (* Error found
   =========================================================================*)
   (*Error Found. Set state to 13, record step and phase number, clear error check flag*)
   IF CCPSystem.Error <> 0 THEN;
   	ErrorCheck := 0;
   	CCPSystem.State := 13;
   	CCPSystem.ErrorStep := PendingStep;
   	CCPSystem.ErrorPhase := PhaseNumber;
   END_IF;
   
   (* No error found
   =========================================================================*)
   (*Complete with no errors. Set state to 0 and clear error check flag*)
   IF PhaseNumber = 5 AND CCPSystem.Error = 0 THEN;
   	ErrorCheck := 0;
   	CCPSystem.State := 0;
   	DTOS (0, CCPSystem.BufferSteps[0]);
   END_IF;
END_ROUTINE

ROUTINE FaultRoutine   (* ladder *)
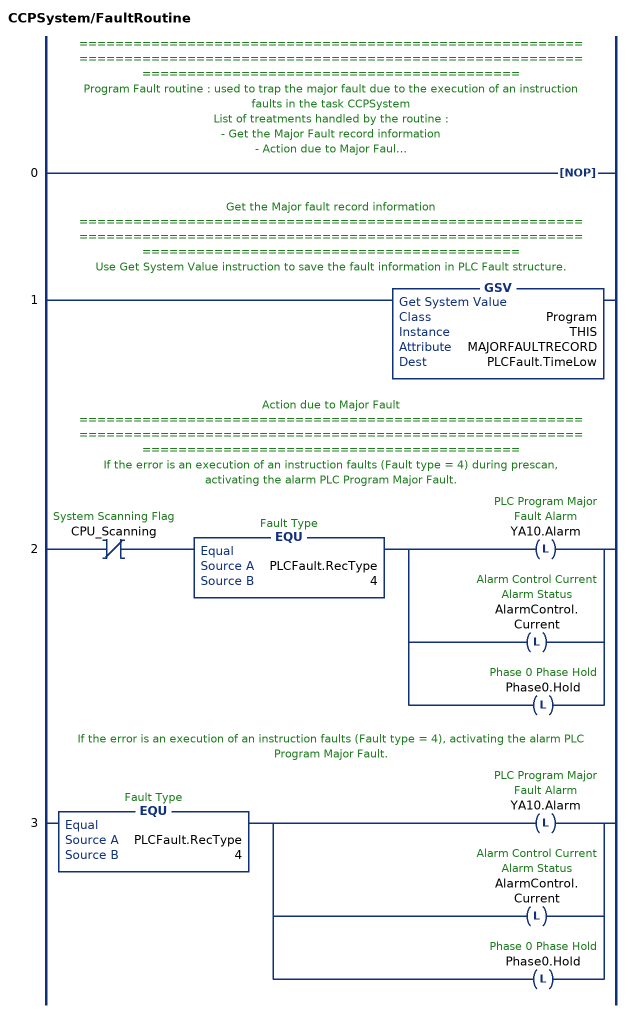
   // ==========================================================================================================================================================
   //                                                            Program Fault routine : used to trap the major fault due to the execution of an instruction faults in the task CCPSystem
   //                                                     List of treatments handled by the routine :
   //                                                          - Get the Major Fault record information
   //                                                          - Action due to Major Fault
   //                                                     -----------------------------------------------------------------------------------------------------------------------------------------------------
   //                                                     History
   // 		2019-DEC-24 - Merck - Q. Spindler - Initial version for Candidate Release 1.00.00.00.a
   // ==========================================================================================================================================================
   0: NOP();
   // Get the Major fault record information
   // ==========================================================================================================================================================
   // Use Get System Value instruction to save the fault information in PLC Fault structure.
   1: GSV(Program,THIS,MAJORFAULTRECORD,PLCFault.TimeLow);
   // Action due to Major Fault
   // ==========================================================================================================================================================
   // If the error is an execution of an instruction faults (Fault type = 4) during prescan, activating the alarm PLC Program Major Fault.
   2: XIO(CPU_Scanning)EQU(PLCFault.RecType,4)[OTL(YA10.Alarm) ,OTL(AlarmControl.Current) ,OTL(Phase0.Hold) ];
   // If the error is an execution of an instruction faults (Fault type = 4), activating the alarm PLC Program Major Fault.
   3: EQU(PLCFault.RecType,4)[OTL(YA10.Alarm) ,OTL(AlarmControl.Current) ,OTL(Phase0.Hold) ];
END_ROUTINE

ROUTINE MainRoutine   (* ladder *)
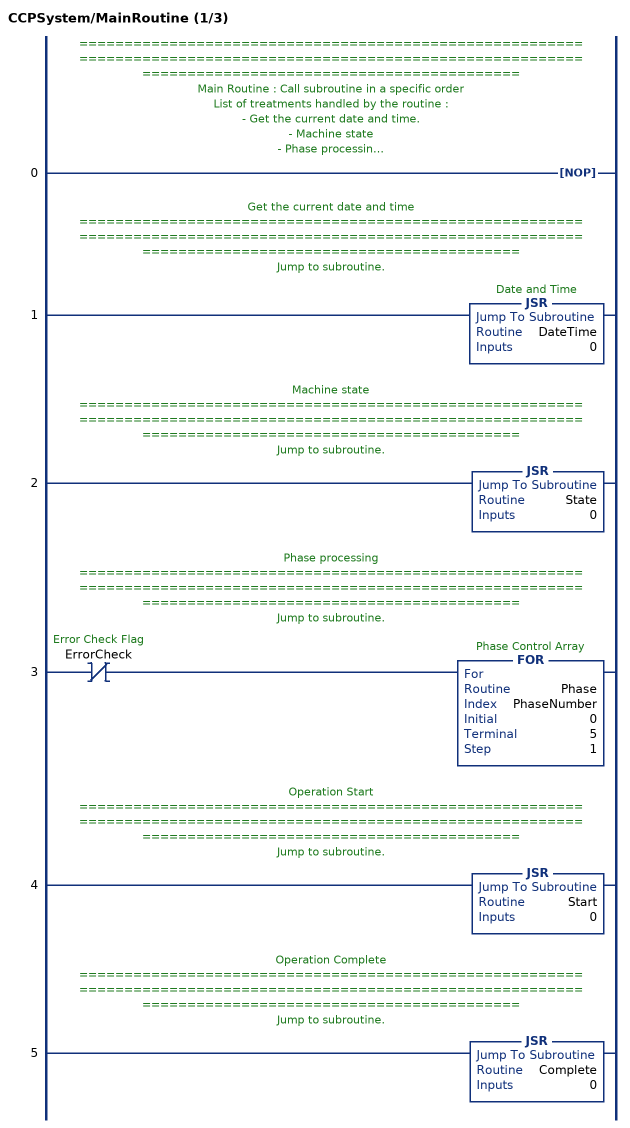
   // ==========================================================================================================================================================
   //                                                                                                            Main Routine : Call subroutine in a specific order
   //                                                     List of treatments handled by the routine :
   //                                                          - Get the current date and time.
   //                                                          - Machine state
   //                                                          - Phase processing
   //                                                          - Operation Start
   //                                                          - Operation Complete
   //                                                          - Procedure timer and totalizer - Hold timer
   //                                                          - Event Log
   //                                                          - CCP System watchdog
   //                                                     -----------------------------------------------------------------------------------------------------------------------------------------------------
   //                                                     History
   // 		2019-DEC-24 - Merck - Q. Spindler - Initial version for Candidate Release 1.00.00.00.a
   //                           2022-JAN-11 - Merck - Q. Spindler - Modifications for Candidate Release 1.01.00.00.a
   // - Add transfer totalizer
   // ========================================================================================================================================================
   0: NOP();
   // Get the current date and time
   // ==========================================================================================================================================================
   // Jump to subroutine.
   1: JSR(DateTime,0);
   // Machine state
   // ==========================================================================================================================================================
   // Jump to subroutine.
   2: JSR(State,0);
   // Phase processing
   // ==========================================================================================================================================================
   // Jump to subroutine.
   3: XIO(ErrorCheck)FOR(Phase,PhaseNumber,0,5,1);
   // Operation Start
   // ==========================================================================================================================================================
   // Jump to subroutine.
   4: JSR(Start,0);
   // Operation Complete
   // ==========================================================================================================================================================
   // Jump to subroutine.
   5: JSR(Complete,0);
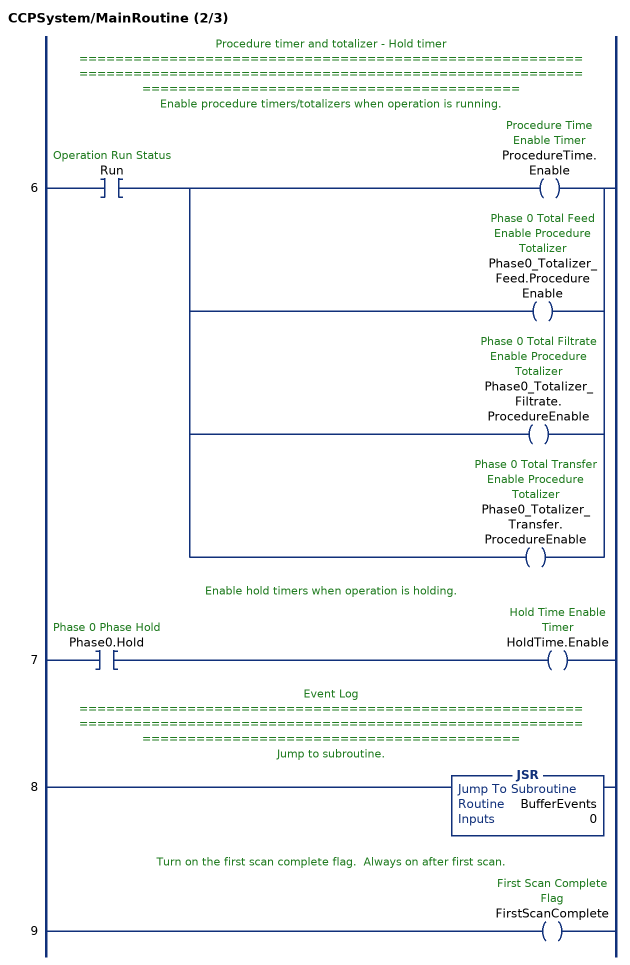
   // Procedure timer and totalizer - Hold timer
   // ==========================================================================================================================================================
   // Enable procedure timers/totalizers when operation is running.
   6: XIC(Run)[OTE(ProcedureTime.Enable) ,OTE(Phase0_Totalizer_Feed.ProcedureEnable) ,OTE(Phase0_Totalizer_Filtrate.ProcedureEnable) ,OTE(Phase0_Totalizer_Transfer.ProcedureEnable) ];
   // Enable hold timers when operation is holding.
   7: XIC(Phase0.Hold)OTE(HoldTime.Enable);
   // Event Log
   // ==========================================================================================================================================================
   // Jump to subroutine.
   8: JSR(BufferEvents,0);
   // Turn on the first scan complete flag.  Always on after first scan.
   9: OTE(FirstScanComplete);
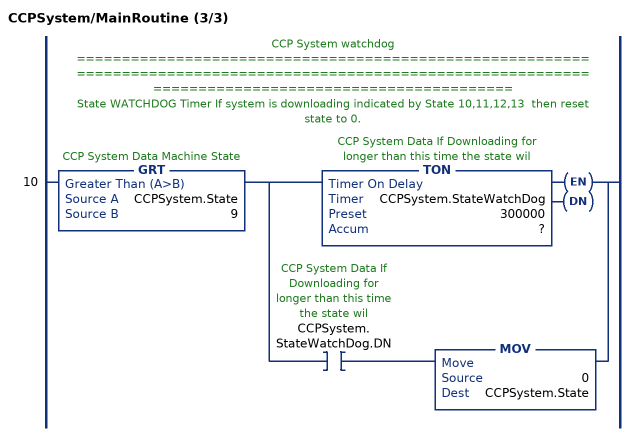
   // CCP System watchdog
   // ==========================================================================================================================================================
   // State WATCHDOG Timer If system is downloading indicated by State 10,11,12,13  then reset state to 0.
   10: GRT(CCPSystem.State,9)[TON(CCPSystem.StateWatchDog,?,?) ,XIC(CCPSystem.StateWatchDog.DN) MOV(0,CCPSystem.State) ];
END_ROUTINE

ROUTINE Phase   (* ladder *)
// Phase Processing Routine
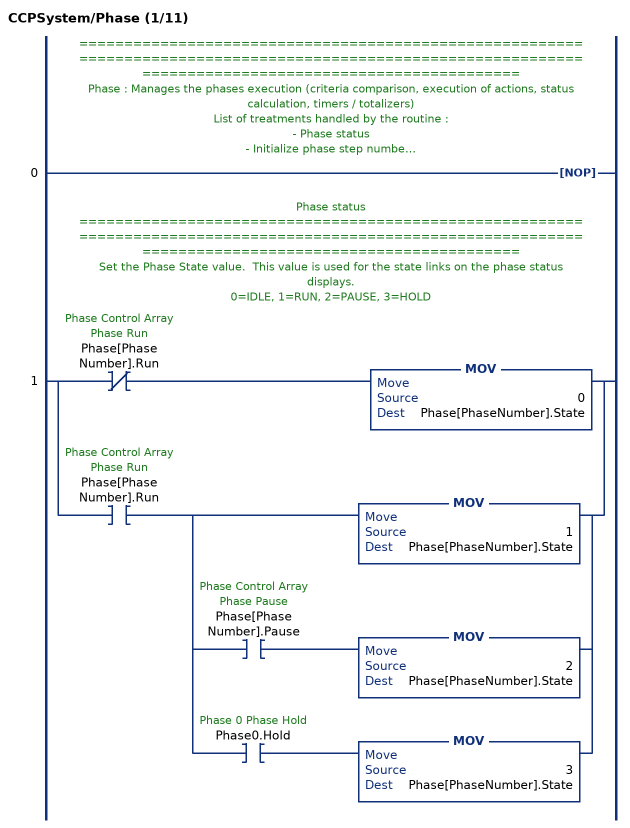
   // ==========================================================================================================================================================
   //                                                                   Phase : Manages the phases execution (criteria comparison, execution of actions, status calculation, timers / totalizers)
   //                                                     List of treatments handled by the routine :
   //                                                          - Phase status
   //                                                          - Initialize phase step number
   //                                                          - Phase Timer / Toalizer
   //                                                          - Phase Stop
   //                                                          - Criteria 1 processing
   //                                                          - Criteria 2 processing
   //                                                          - Jump Step
   //                                                          - Criteria met
   //                                                          - Phase Pause
   //                                                          - Prompt processing
   //                                                          - Branch step processing
   //                                                          - Action processing
   //                                                          - Update step number
   //                                                          - Reset step timer and totalizer
   //                                                     -----------------------------------------------------------------------------------------------------------------------------------------------------
   //                                                     History
   // 		2019-DEC-24 - Merck - Q. Spindler - Initial version for Candidate Release 1.00.00.00.a
   //                                  2020-APR-06 - Merck - Q. Spindler - Modifications for Candidate Release 1.00.00.00.b
   //                                      Replace TimerControl.Tick by TimerControl.TickMainTask
   //                                  2021-APR-22 - Merck - Q. Spindler - Modifications for Candidate Release 1.00.00.00.e
   //                                     - Add Reset of crit1metTime when the totalizers are reset
   //                           2022-JAN-11 - Merck - Q. Spindler - Modifications for Candidate Release 1.01.00.00.a
   // - Add transfer totalizer
   //                           2022-SEP-20 - Actemium - J. Jaekel - Modifications for Candidate Release 1.01.00.01.a
   // - Add Hold condition for Criteria 1 met timer
   // ========================================================================================================================================================
   0: NOP();
   // Phase status
   // ==========================================================================================================================================================
   // Set the Phase State value.  This value is used for the state links on the phase status displays.
   // 0=IDLE, 1=RUN, 2=PAUSE, 3=HOLD
   1: [XIO(Phase[PhaseNumber].Run) MOV(0,Phase[PhaseNumber].State) ,XIC(Phase[PhaseNumber].Run) [MOV(1,Phase[PhaseNumber].State) ,XIC(Phase[PhaseNumber].Pause) MOV(2,Phase[PhaseNumber].State) ,XIC(Phase0.Hold) MOV(3,Phase[PhaseNumber].State) ] ];
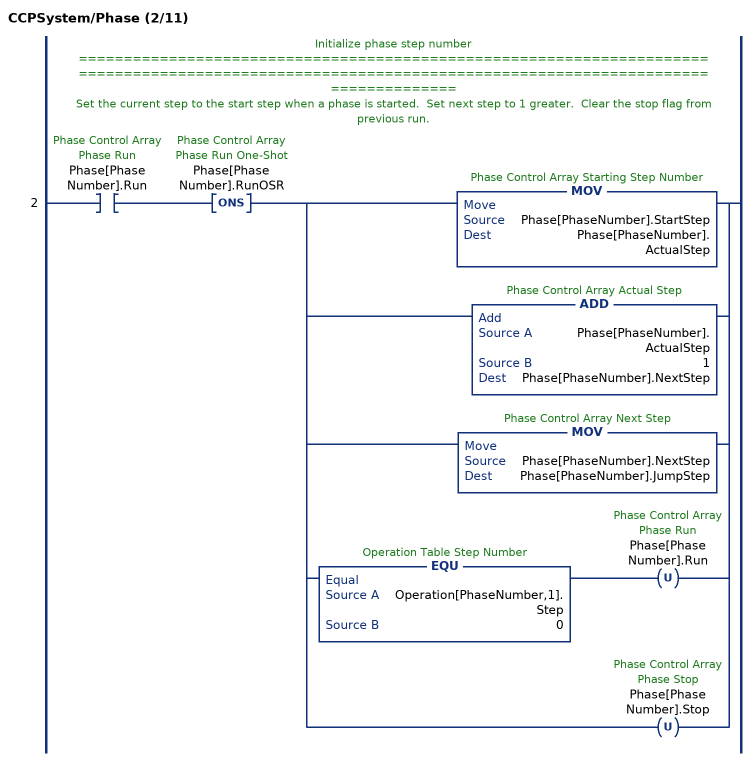
   // Initialize phase step number
   // ==========================================================================================================================================================
   // Set the current step to the start step when a phase is started.  Set next step to 1 greater.  Clear the stop flag from previous run.
   2: XIC(Phase[PhaseNumber].Run)ONS(Phase[PhaseNumber].RunOSR)[MOV(Phase[PhaseNumber].StartStep,Phase[PhaseNumber].ActualStep) ,ADD(Phase[PhaseNumber].ActualStep,1,Phase[PhaseNumber].NextStep) ,MOV(Phase[PhaseNumber].NextStep,Phase[PhaseNumber].JumpStep) ,EQU(Operation[PhaseNumber,1].Step,0) OTU(Phase[PhaseNumber].Run) ,OTU(Phase[PhaseNumber].Stop) ];
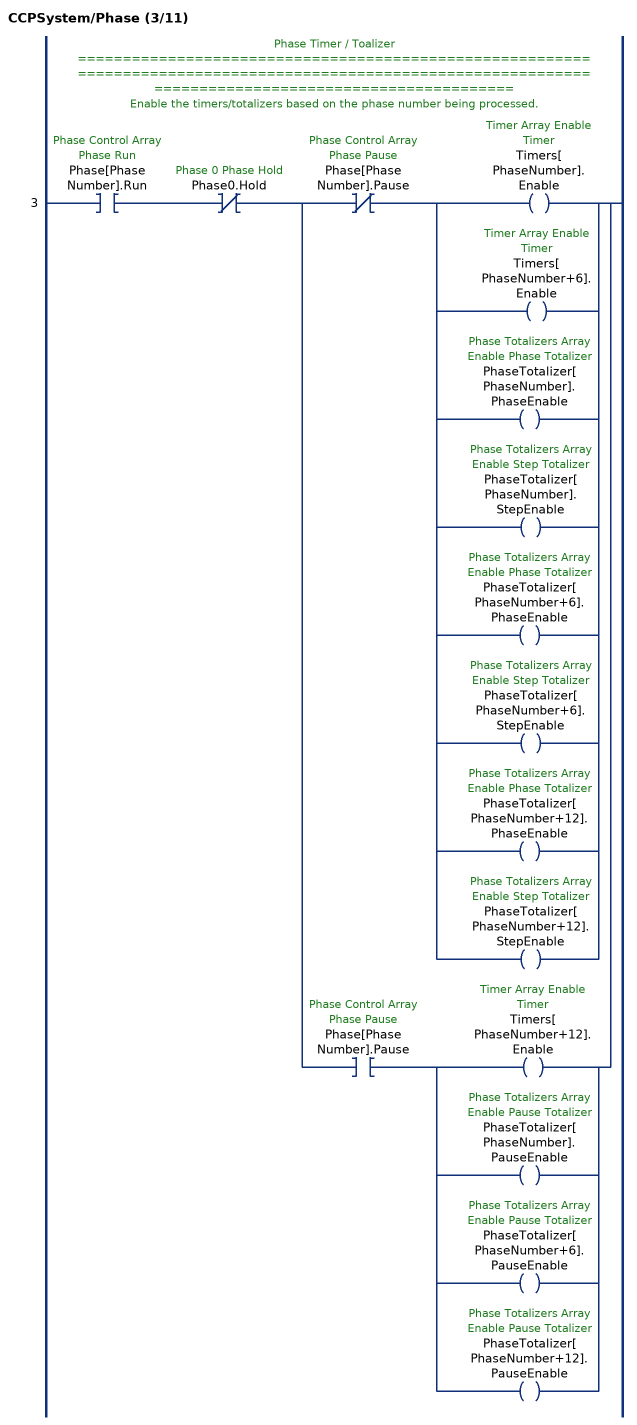
   // Phase Timer / Toalizer
   // ==========================================================================================================================================================
   // Enable the timers/totalizers based on the phase number being processed.
   3: XIC(Phase[PhaseNumber].Run)XIO(Phase0.Hold)[XIO(Phase[PhaseNumber].Pause) [OTE(Timers[PhaseNumber].Enable) ,OTE(Timers[PhaseNumber+6].Enable) ,OTE(PhaseTotalizer[PhaseNumber].PhaseEnable) ,OTE(PhaseTotalizer[PhaseNumber].StepEnable) ,OTE(PhaseTotalizer[PhaseNumber+6].PhaseEnable) ,OTE(PhaseTotalizer[PhaseNumber+6].StepEnable) ,OTE(PhaseTotalizer[PhaseNumber+12].PhaseEnable) ,OTE(PhaseTotalizer[PhaseNumber+12].StepEnable) ] ,XIC(Phase[PhaseNumber].Pause) [OTE(Timers[PhaseNumber+12].Enable) ,OTE(PhaseTotalizer[PhaseNumber].PauseEnable) ,OTE(PhaseTotalizer[PhaseNumber+6].PauseEnable) ,OTE(PhaseTotalizer[PhaseNumber+12].PauseEnable) ] ];
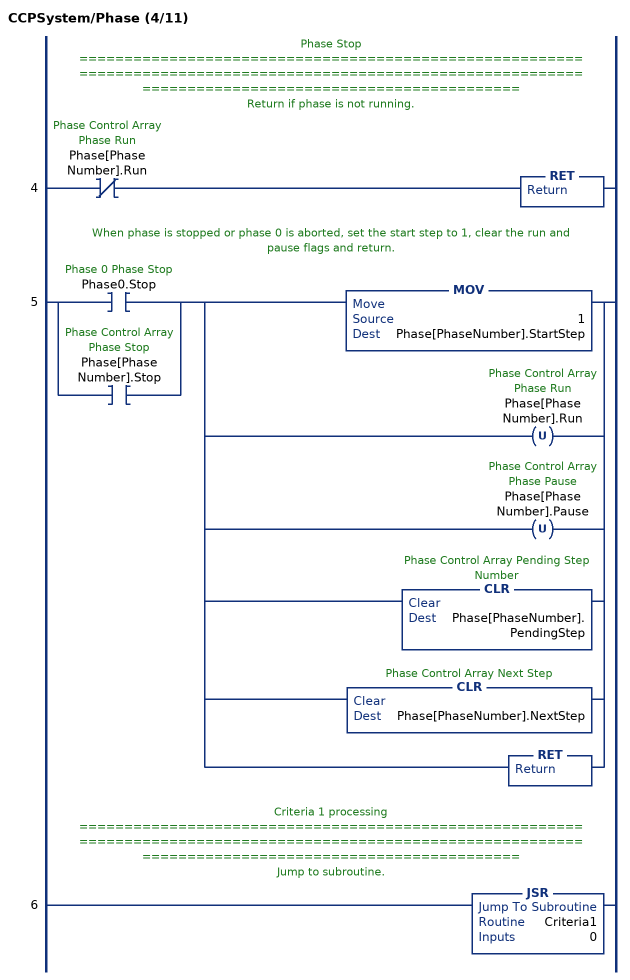
   // Phase Stop
   // ==========================================================================================================================================================
   // Return if phase is not running.
   4: XIO(Phase[PhaseNumber].Run)RET();
   // When phase is stopped or phase 0 is aborted, set the start step to 1, clear the run and pause flags and return.
   5: [XIC(Phase0.Stop) ,XIC(Phase[PhaseNumber].Stop) ][MOV(1,Phase[PhaseNumber].StartStep) ,OTU(Phase[PhaseNumber].Run) ,OTU(Phase[PhaseNumber].Pause) ,CLR(Phase[PhaseNumber].PendingStep) ,CLR(Phase[PhaseNumber].NextStep) ,RET() ];
   // Criteria 1 processing
   // ==========================================================================================================================================================
   // Jump to subroutine.
   6: JSR(Criteria1,0);
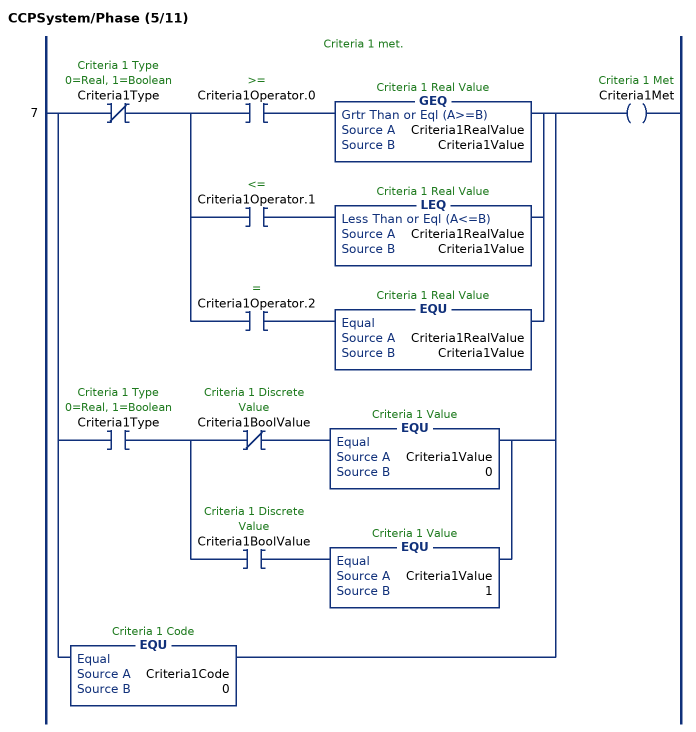
   // Criteria 1 met.
   7: [XIO(Criteria1Type) [XIC(Criteria1Operator.0) GEQ(Criteria1RealValue,Criteria1Value) ,XIC(Criteria1Operator.1) LEQ(Criteria1RealValue,Criteria1Value) ,XIC(Criteria1Operator.2) EQU(Criteria1RealValue,Criteria1Value) ] ,XIC(Criteria1Type) [XIO(Criteria1BoolValue) EQU(Criteria1Value,0) ,XIC(Criteria1BoolValue) EQU(Criteria1Value,1) ] ,EQU(Criteria1Code,0) ]OTE(Criteria1Met);
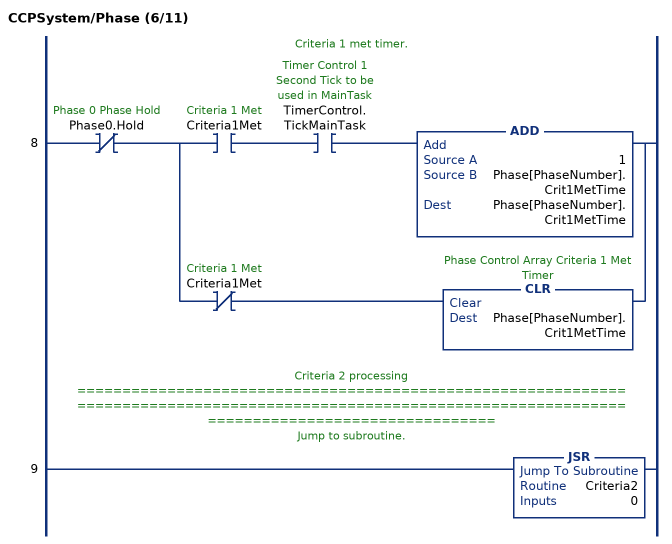
   // Criteria 1 met timer.
   8: XIO(Phase0.Hold)[XIC(Criteria1Met) XIC(TimerControl.TickMainTask) ADD(1,Phase[PhaseNumber].Crit1MetTime,Phase[PhaseNumber].Crit1MetTime) ,XIO(Criteria1Met) CLR(Phase[PhaseNumber].Crit1MetTime) ];
   // Criteria 2 processing
   // ==========================================================================================================================================================
   // Jump to subroutine.
   9: JSR(Criteria2,0);
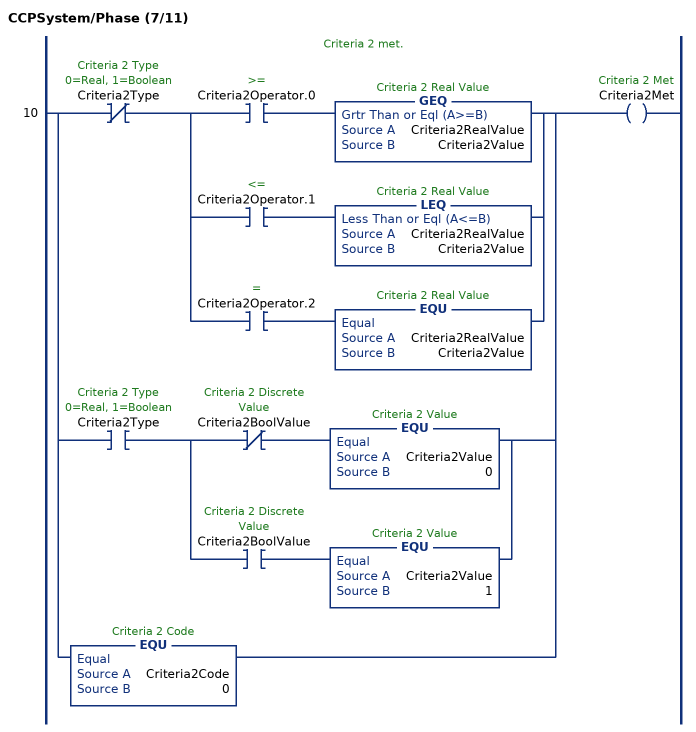
   // Criteria 2 met.
   10: [XIO(Criteria2Type) [XIC(Criteria2Operator.0) GEQ(Criteria2RealValue,Criteria2Value) ,XIC(Criteria2Operator.1) LEQ(Criteria2RealValue,Criteria2Value) ,XIC(Criteria2Operator.2) EQU(Criteria2RealValue,Criteria2Value) ] ,XIC(Criteria2Type) [XIO(Criteria2BoolValue) EQU(Criteria2Value,0) ,XIC(Criteria2BoolValue) EQU(Criteria2Value,1) ] ,EQU(Criteria2Code,0) ]OTE(Criteria2Met);
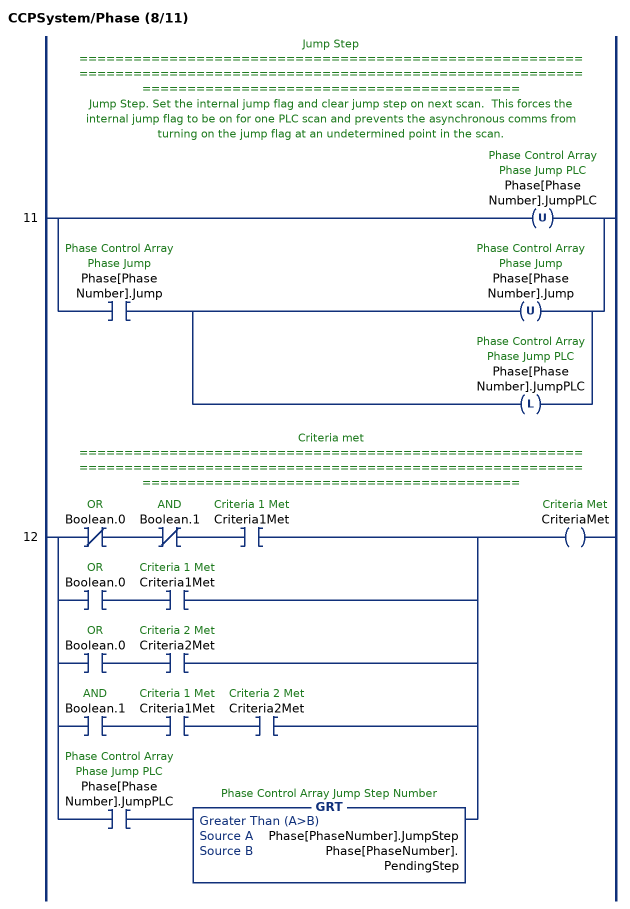
   // Jump Step
   // ==========================================================================================================================================================
   // Jump Step. Set the internal jump flag and clear jump step on next scan.  This forces the internal jump flag to be on for one PLC scan and prevents the asynchronous comms from turning on the jump flag at an undetermined point in the scan.
   11: [OTU(Phase[PhaseNumber].JumpPLC) ,XIC(Phase[PhaseNumber].Jump) [OTU(Phase[PhaseNumber].Jump) ,OTL(Phase[PhaseNumber].JumpPLC) ] ];
   // Criteria met
   // ==========================================================================================================================================================
   12: [XIO(Boolean.0) XIO(Boolean.1) XIC(Criteria1Met) ,XIC(Boolean.0) XIC(Criteria1Met) ,XIC(Boolean.0) XIC(Criteria2Met) ,XIC(Boolean.1) XIC(Criteria1Met) XIC(Criteria2Met) ,XIC(Phase[PhaseNumber].JumpPLC) GRT(Phase[PhaseNumber].JumpStep,Phase[PhaseNumber].PendingStep) ]OTE(CriteriaMet);
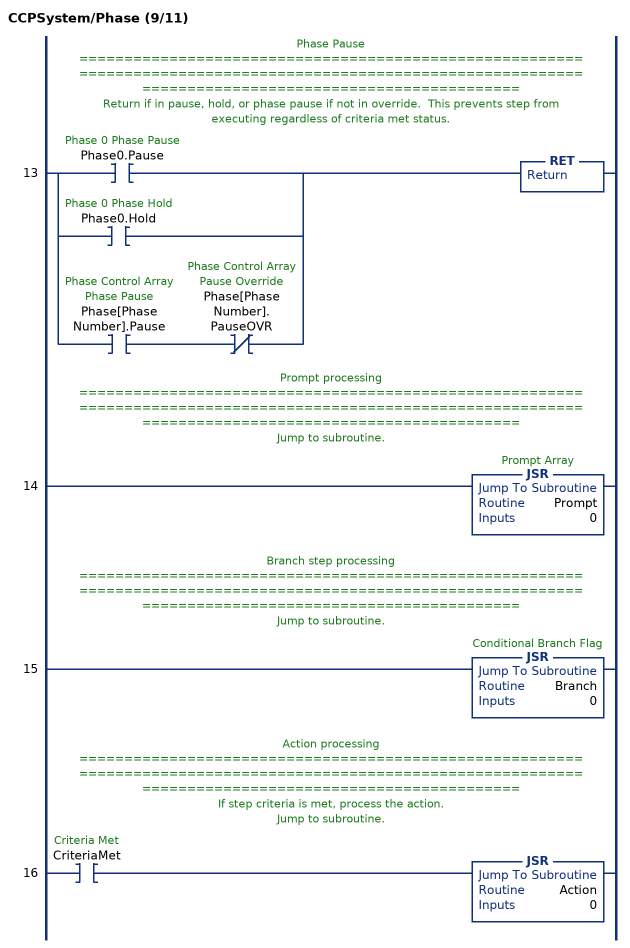
   // Phase Pause
   // ==========================================================================================================================================================
   // Return if in pause, hold, or phase pause if not in override.  This prevents step from executing regardless of criteria met status.
   13: [XIC(Phase0.Pause) ,XIC(Phase0.Hold) ,XIC(Phase[PhaseNumber].Pause) XIO(Phase[PhaseNumber].PauseOVR) ]RET();
   // Prompt processing
   // ==========================================================================================================================================================
   // Jump to subroutine.
   14: JSR(Prompt,0);
   // Branch step processing
   // ==========================================================================================================================================================
   // Jump to subroutine.
   15: JSR(Branch,0);
   // Action processing
   // ==========================================================================================================================================================
   // If step criteria is met, process the action.
   // Jump to subroutine.
   16: XIC(CriteriaMet)JSR(Action,0);
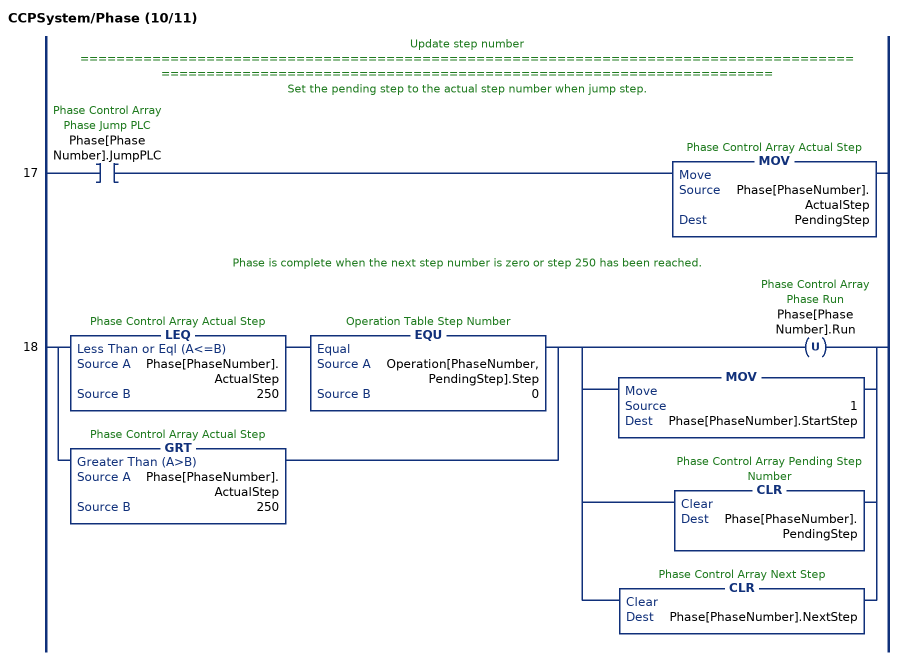
   // Update step number
   // ==========================================================================================================================================================
   // Set the pending step to the actual step number when jump step.
   17: XIC(Phase[PhaseNumber].JumpPLC)MOV(Phase[PhaseNumber].ActualStep,PendingStep);
   // Phase is complete when the next step number is zero or step 250 has been reached.
   18: [LEQ(Phase[PhaseNumber].ActualStep,250) EQU(Operation[PhaseNumber,PendingStep].Step,0) ,GRT(Phase[PhaseNumber].ActualStep,250) ][OTU(Phase[PhaseNumber].Run) ,MOV(1,Phase[PhaseNumber].StartStep) ,CLR(Phase[PhaseNumber].PendingStep) ,CLR(Phase[PhaseNumber].NextStep) ];
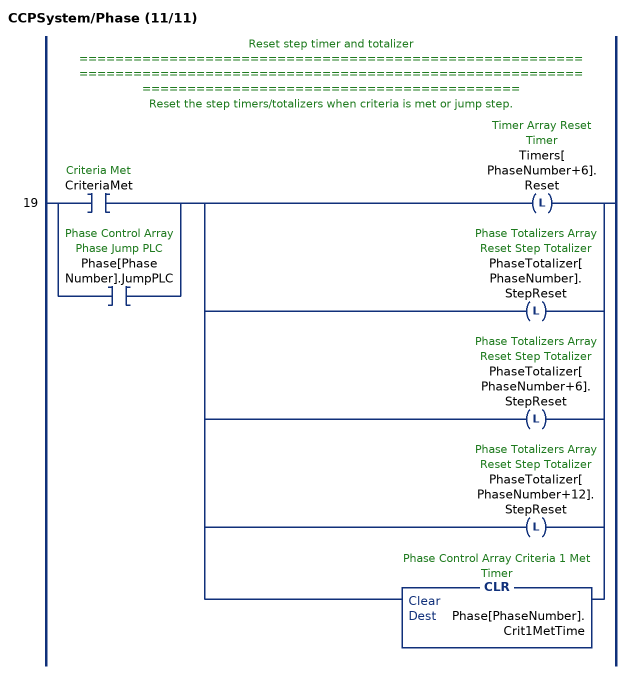
   // Reset step timer and totalizer
   // ==========================================================================================================================================================
   // Reset the step timers/totalizers when criteria is met or jump step.
   19: [XIC(CriteriaMet) ,XIC(Phase[PhaseNumber].JumpPLC) ][OTL(Timers[PhaseNumber+6].Reset) ,OTL(PhaseTotalizer[PhaseNumber].StepReset) ,OTL(PhaseTotalizer[PhaseNumber+6].StepReset) ,OTL(PhaseTotalizer[PhaseNumber+12].StepReset) ,CLR(Phase[PhaseNumber].Crit1MetTime) ];
END_ROUTINE
